// TwinCAT 3 PLC project PLC1
// ProgramVersion: 3.1.4024.0
// libraries:
//   Tc2_MC2, * (Beckhoff Automation GmbH)
//   Tc2_Standard, * (Beckhoff Automation GmbH)
//   Tc2_System, * (Beckhoff Automation GmbH)
//   Tc2_TcpIp, * (Beckhoff Automation GmbH)
//   Tc3_Module, * (Beckhoff Automation GmbH)
// project tree:
//   DUTs/ E_MelsecDevice.TcDUT, ST_MelsecSession.TcDUT, ST_QueuedCameraProduct.TcDUT, ST_Point2D.TcDUT, ST_QD75_Command.TcDUT, ST_QD75_Feedback.TcDUT
//   GVLs/ GVL_MD200_IO.TcGVL, GVL.TcGVL
//   / PlcTask.TcTTO
//   POUs/ FB_ConveyorEncoder.TcPOU, FB_ConveyorTracking4Pt.TcPOU, FB_InovanceMD200Conveyor.TcPOU, FB_EziServoControl.TcPOU, FB_MelsecEchoVerify.TcPOU, FB_MelsecDebugXY4Pt.TcPOU, FB_CameraProductQueue.TcPOU, FB_UpstreamCameraTracking4Pt.TcPOU, FB_XYTrackingManualAck.TcPOU, FB_MelsecRead.TcPOU, FB_MelsecTcpConfig.TcPOU, FB_MelsecWrite.TcPOU, FB_QD75CommandPublisher.TcPOU, MAIN.TcPOU
// real-time tasks:
//   TASK PlcTask: cycle T#10ms, priority 20, ADS port 350
// motion (NC):
//   TASK NC-Task 1 SAF: cycle T#2ms, priority 4, ADS port 501
//   TASK NC-Task 1 SVB: cycle T#10ms, priority 8, ADS port 511
//   AXIS Axis 1 (id 2)
//     General: UnitName=Degree
//     Velo: Maximum=50000
//     OtherSettings: AllowMotionCmdToSlave=true
//     encoder EncType=19
//       EncPara: ScaleFactorNumerator=360, ScaleFactorDenominator=10000, MaxCount=#xffffffff
//     drive DrvType=16
//       DrvPara: MaxCount=#xffffffff, DriveControlDWord=#x00020000
//         Analog: VeloReferenz=60000, TorqueSetpointScale=10, ScaleFactorActTorque=0.1
//         TimeComp: TaskDelayCycles=1
//     controller CtrType=1
//       CtrPara: PriorControlFactor=1
//         PosDiffControl: Range=60, Time=0.05
//         Observer: BandWidth=20
// I/O:
//   DEVICE Device 2 (EtherCAT), AmsNetId 10.81.27.140.3.1
//     Box 1 (NA-9286,Crevis) [NA-9286 EtherCAT Adapter, Crevis]
//       modules: Module 1 (ST-5101), Module 2 (ST-1228), Module 3 (ST-1228), Module 4 (ST-1228), Module 5 (ST-1228), Module 6 (ST-1228), Module 7 (ST-2318), Module 8 (ST-2318), Module 9 (ST-2318), Module 10 (ST-2318), Module 11 (ST-4424), Module 12 (ST-5114), Module 13 (ST-3214)
//     Drive 2 (Ezi-SERVO2 EtherCAT) [Ezi-SERVO2 EtherCAT]
// variable links:
//   NC-Task 1 SAF/Axes/Axis 1 <-> Device 2 (EtherCAT)/Drive 2 (Ezi-SERVO2 EtherCAT)
//     Drive/Inputs/In/nDcOutputTime <-> InfoData/DcOutputShift
//     Drive/Inputs/In/nState1 <-> CSP Inputs/Status Word
//     Drive/Inputs/In/nState2 <-> CSP Inputs/Status Word @bit 8
//     Drive/Inputs/In/nState4 @bit 1 <-> WcState/InputToggle
//     Drive/Inputs/In/nState4 <-> WcState/WcState
//     Drive/Outputs/Out/nCtrl1 <-> CSP Outputs/Control Word
//     Drive/Outputs/Out/nCtrl2 <-> CSP Outputs/Control Word @bit 8
//     Drive/Outputs/Out/nDataOut1 <-> CSP Outputs/Target Position
//     Enc/Inputs/In/nDataIn1 <-> CSP Inputs/Position Actual Value
//     Enc/Inputs/In/nDataIn3 <-> CSP Inputs/Touch probe 1 positive value
//     Enc/Inputs/In/nDataIn5 <-> CSP Inputs/Touch probe 2 positive value
//     Enc/Inputs/In/nDcInputTime <-> InfoData/DcInputShift
//     Enc/Inputs/In/nState4 @bit 1 <-> WcState/InputToggle
//     Enc/Inputs/In/nState4 <-> WcState/WcState
//     Enc/Inputs/In/nState5 <-> CSP Inputs/Touch probe status
//     Enc/Inputs/In/nState6 <-> CSP Inputs/Touch probe status @bit 8
//     Enc/Outputs/Out/nCtrl5 <-> CSP Outputs/Touch probe function
//     Enc/Outputs/Out/nCtrl6 <-> CSP Outputs/Touch probe function @bit 8
//   PLC1/PLC1 Instance <-> Device 2 (EtherCAT)/Box 1 (NA-9286,Crevis)
//     PlcTask Inputs/GVL.aIn[{0..15}] <-> Module 12 (ST-5114)/Input(s)/Byte {0..15}  (16 links)
//     PlcTask Inputs/GVL_MD200_IO.bEStopFeedback <-> Module 6 (ST-1228)/Input(s)/Byte 0
//     PlcTask Outputs/GVL.aOut[{0..3}] <-> Module 12 (ST-5114)/Output(s)/Byte {0..3}  (4 links)
//     PlcTask Outputs/GVL_MD200_IO.bRUN_DO <-> Module 10 (ST-2318)/Output(s)/Byte 0
//     PlcTask Outputs/GVL_MD200_IO.nAO1_Raw <-> Module 11 (ST-4424)/Output(s)/Analog Output Ch#1 Byte
//   PLC1/PLC1 Instance <-> NC-Task 1 SAF/Axes/Axis 1
//     PlcTask Inputs/MAIN.Axis1.NcToPlc <-> Outputs/ToPlc
//     PlcTask Outputs/MAIN.Axis1.PlcToNc <-> Inputs/FromPlc

CONFIGURATION PLC1
    RESOURCE PLC ON TwinCAT3
        TASK PlcTask(INTERVAL := T#10ms, PRIORITY := 20);
        PROGRAM MAIN WITH PlcTask : MAIN;
    END_RESOURCE
END_CONFIGURATION

// ---- DUTs/E_MelsecDevice.TcDUT
// Mã định danh vùng nhớ phần cứng Mitsubishi theo chuẩn MC Protocol Binary 3E Frame
TYPE E_MelsecDevice :
(
    DEV_D   := 16#A8, // Thanh ghi dữ liệu D (Data Register) - Word
    DEV_M   := 16#90, // Rơ-le nội bộ M (Internal Relay) - Bit / Word
    DEV_W   := 16#B4, // Thanh ghi liên kết W (Link Register) - Word
    DEV_R   := 16#AF, // Thanh ghi tệp R (File Register) - Word
    DEV_ZR  := 16#B0, // Thanh ghi tệp liên tục ZR (File Register Consecutive) - Word
    DEV_X   := 16#9C, // Ngõ vào vật lý X (Input) - Bit
    DEV_Y   := 16#9D, // Ngõ ra vật lý Y (Output) - Bit
    DEV_B   := 16#A0, // Rơ-le liên kết B (Link Relay) - Bit / Word
    DEV_L   := 16#92, // Rơ-le chốt L (Latch Relay) - Bit
    DEV_TN  := 16#C2, // Giá trị hiện tại Timer TN (Timer Current Value) - Word
    DEV_CN  := 16#C5  // Giá trị hiện tại Counter CN (Counter Current Value) - Word
);
END_TYPE

// ---- DUTs/ST_MelsecSession.TcDUT
TYPE ST_MelsecSession :
STRUCT
    hSocket     : T_HSOCKET; // Socket TCP dùng chung
    bConnected  : BOOL;      // TRUE khi đã kết nối PLC
    bBusy       : BOOL;      // TRUE khi Read hoặc Write đang giao dịch
    bError      : BOOL;      // Lỗi cuối cùng
    nErrorID    : UDINT;     // Mã lỗi cuối cùng
END_STRUCT
END_TYPE

// ---- DUTs/ST_QueuedCameraProduct.TcDUT
TYPE ST_QueuedCameraProduct :
STRUCT
    bValid                    : BOOL;
    nProductID                : UDINT;
    nState                    : INT; // 0 EMPTY, 1 WAIT_ROBOT, 2 GEOMETRIC_WINDOW
    bAllCornersInside         : BOOL;
    bForecastWindowOK         : BOOL;
    rEncoderAtExposure_mm     : LREAL;
    rCenterAtExposureX_mm     : LREAL;
    rCenterAtExposureY_mm     : LREAL;
    rThetaRobot_deg           : LREAL;
    rTravel_mm                : LREAL;
    rCenterNowX_mm            : LREAL;
    rCenterNowY_mm            : LREAL;
    aCornerBase               : ARRAY[1..4] OF ST_Point2D;
    aCornerNow                : ARRAY[1..4] OF ST_Point2D;
END_STRUCT
END_TYPE

// ---- DUTs/ST_Point2D.TcDUT
TYPE ST_Point2D :
STRUCT
    X : LREAL; // Tọa độ X (mm)
    Y : LREAL; // Tọa độ Y (mm)
END_STRUCT
END_TYPE

// ---- DUTs/ST_QD75_Command.TcDUT
TYPE ST_QD75_Command :
STRUCT
    Target_X       : DINT; // D100..D101: Tọa độ đón đầu trục X (0.1 um)
    Target_Y       : DINT; // D102..D103: Tọa độ trục Y đỉnh (0.1 um)
    Target_Z_Down  : DINT; // D104..D105: Độ cao hạ chấm keo (0.1 um, 4.0mm = 40000)
    Speed_Approach : DINT; // D106..D107: Vận tốc bay nội suy 3 trục (0.01 mm/min, 500mm/s = 3000000)
    Speed_Sync     : DINT; // D108..D109: Vận tốc đồng tốc trục X khi chấm keo (= V_conv * 6000)
    DeltaX_Sync    : DINT; // D110..D111: Quãng đường trượt đồng tốc 60ms (0.1 um)
    Target_Z_Safe  : DINT; // D112..D113: Độ cao an toàn khi rút kim (0.1 um, 0.0mm = 0)
    Vertex_Index   : INT;  // D114: Thứ tự đỉnh đang làm (1..4)
    Cmd_Start      : BOOL; // M1000: Kích chạy đỉnh đang nạp (TwinCAT -> PLC-Q)
END_STRUCT
END_TYPE

// ---- DUTs/ST_QD75_Feedback.TcDUT
TYPE ST_QD75_Feedback :
STRUCT
    Ack_Done    : BOOL; // M1001: PLC-Q báo Point 3 hoàn tất
    Robot_Busy  : BOOL; // M102: PLC-Q đang kiểm tra/nạp/chạy
    In_Position : BOOL; // M103: Đỉnh đã hoàn tất, chờ Master hạ M1000
    Robot_Alarm : BOOL; // M104: QD75 hoặc kiểm tra biên báo lỗi
END_STRUCT
END_TYPE

// ---- GVLs/GVL_MD200_IO.TcGVL
VAR_GLOBAL
    // E-stop circuit HEALTHY auxiliary contact feedback.
    // REVIEW BEFORE ACTIVATION: maps ST-1228 SLOT 6 / DI0 (physical terminal 0).
    // This is a PROPOSED wiring channel, not confirmed by cabinet visual inspection.
    // It must be wired to the healthy auxiliary feedback of an independent
    // hardwired emergency-stop safety circuit. TRUE = safety chain healthy.
    // This input alone is NOT an emergency-stop device.
    {attribute 'TcLinkToOSO' := '<0,1,0>TIID^Device 2 (EtherCAT)^Box 1 (NA-9286,Crevis)^Module 6 (ST-1228)^Input(s)^Byte 0'}
    bEStopFeedback AT %I* : BOOL := FALSE;

    // MD200 physical process-image channels, staged for deliberate link review.
    // ST-4424 Module 11 Channel AO1 (physical terminal 1, 0-10V).
    // UINT 16 bit with 12-bit useful range 0..4095.
    {attribute 'TcLinkTo' := 'TIID^Device 2 (EtherCAT)^Box 1 (NA-9286,Crevis)^Module 11 (ST-4424)^Output(s)^Analog Output Ch#1 Byte'}
    nAO1_Raw AT %Q* : UINT := 0;

    // Staged logical RUN: ST-2318 Module 10 immediately before AO module.
    // DO0 is bit 0 of Output(s)^Byte 0; map ONLY one bit (not entire BYTE).
    // WARNING: physical DO0/pin 0 must be confirmed unused and NPN wiring
    // checked by the on-site technician BEFORE activating this configuration.
    // All runtime software permits remain FALSE by default.
    {attribute 'TcLinkToOSO' := '<0,1,0>TIID^Device 2 (EtherCAT)^Box 1 (NA-9286,Crevis)^Module 10 (ST-2318)^Output(s)^Byte 0'}
    bRUN_DO AT %Q* : BOOL := FALSE;
END_VAR

// ---- GVLs/GVL.TcGVL
VAR_GLOBAL
    aIn  AT %I* : ARRAY[0..15] OF BYTE;  // TxPDO 16 byte
    aOut AT %Q* : ARRAY[0..3]  OF BYTE;  // RxPDO 4 byte
END_VAR

// ---- POUs/MAIN.TcPOU
PROGRAM MAIN
VAR
    // ================================================================
    // 1. KẾT NỐI TCP VỚI CPU MITSUBISHI Q06UDEH (CỔNG 5010)
    // ================================================================
    stMelsec            : ST_MelsecSession; // Session TCP dùng chung
    fbMelsecConfig      : FB_MelsecTcpConfig;

    bTcpEnable          : BOOL := TRUE;     // Tự động kết nối và duy trì kết nối mạng
    sPlcQ_IP            : STRING(15) := '192.168.3.39'; // IP của PLC-Q
    nPlcQ_Port          : UDINT := 5010;   // Cổng Port MC Protocol 5010

    bPlcQConnected      : BOOL;             // ĐÈN BÁO: TRUE = Đã thông mạng với PLC-Q
    bPlcQError          : BOOL;
    nPlcQErrorID        : UDINT;

    // ================================================================
    // 2. TEST TRUYỀN THÔNG THỦ CÔNG SANG PLC-Q (KHI bStartGlueCycle = FALSE)
    // ================================================================
    bTest_WriteD100     : BOOL := FALSE;    // Click đúp TRUE -> Ghi nTest_D100_Val vào D100-D101
    nTest_D100_Val      : DINT := 100;      // Số 32-bit gửi thử sang D100
    bTest_WriteM1000    : BOOL := FALSE;    // Click đúp TRUE -> Ghi bit M1000
    bTest_M1000_Val     : BOOL := TRUE;     // Giá trị bit M1000 muốn ghi (TRUE=ON, FALSE=OFF)
    bTest_ReadM1001     : BOOL := FALSE;    // Click đúp TRUE -> Đọc bit M1001 từ PLC-Q
    bTest_M1001_Result  : BOOL;             // Giá trị M1001 đọc được từ PLC-Q

    // ================================================================
    // 3. ENCODER BĂNG TẢI: ST-5114 MODULE 12
    // ================================================================
    fbConveyor          : FB_ConveyorEncoder;

    nEncoderPulse       : UINT;            // HARDWARE RAW counter, NOT zeroed on TwinCAT boot
    nEncoderPulseSinceStart : DINT := 0; // VIRTUAL count starting from 0 on PLC boot
    nEncoderDelta       : INT;             // Xung thay đổi trong 10 ms
    rConveyorSpeed      : LREAL;           // Vận tốc băng tải lọc mượt, mm/s
    rConveyorSpeedMPM   : LREAL;           // Vận tốc băng tải, m/phút
    rConveyorDist       : LREAL;           // Tổng quãng đường băng tải, mm

    // ================================================================
    // ================================================================
    // MD200 VFD PREPARATION / VIRTUAL ONLY (NO PHYSICAL I/O MAPPING).
    // Outputs remain disconnected from Crevis ST-2318 and ST-4424.
    // ================================================================
    fbMD200_VFD               : FB_InovanceMD200Conveyor;
    // Global normal-PLC motion inhibit, NOT an emergency stop safety function.
    // TRUE only when the auxiliary feedback from hardwired EStop is healthy.
    bSystemEStopOK             : BOOL := FALSE;
    bSystemStopRequested       : BOOL := TRUE;
    // Only 3 operator-visible MD200 signals: EStopOK monitor, START and Hz.
    // EStopOK is derived from the wired digital feedback, NOT an HMI override.
    bMD200_EStopOK           : BOOL := FALSE;
    bMD200_Start             : BOOL := FALSE;
    rMD200_SetFrequency_Hz    : LREAL := 0.0;
    // Diagnostics (read-only outputs from the FB)
    bMD200_DO_RunVirtual      : BOOL;
    nMD200_AO_RawVirtual      : INT;
    rMD200_AO_VoltsVirtual    : LREAL;
    rMD200_Target_Hz          : LREAL;
    rMD200_Ramped_Hz          : LREAL;
    bMD200_AtTarget           : BOOL;
    bMD200_Limited            : BOOL;
    nMD200_Status             : UINT;

    // ================================================================
    // 4. EZI-SERVO: TRỤC QUAY ĐƠN VỊ DEGREE
    // ================================================================
    Axis1               : AXIS_REF;

    fbServo             : FB_EziServoControl;

    bServo_Enable       : BOOL := FALSE;     // TRUE = Servo ON / giữ cốt
    bServo_Reset        : BOOL := FALSE;    // TRUE một chu kỳ = Reset Alarm
    bServo_JogFwd       : BOOL := FALSE;    // TRUE = chạy thuận
    bServo_JogBwd       : BOOL := FALSE;    // TRUE = chạy nghịch

    rServo_Speed        : LREAL := 100.0;   // Degree/s
    rServo_Acc          : LREAL := 400.0;   // Degree/s2
    rServo_Dec          : LREAL := 400.0;   // Degree/s2

    bServo_Ready        : BOOL;             // TRUE = Servo ON
    rServo_ActPos_Deg   : LREAL;            // Góc thực tế, Degree
    rServo_ActVel_Deg_s : LREAL;            // Vận tốc thực tế, Degree/s

    // ================================================================
    // 5. TRACKING 4 ĐIỂM: CAMERA + ENCODER
    // ================================================================
    fbTracking4Pt       : FB_ConveyorTracking4Pt;

    bSystemReset        : BOOL := FALSE;    // TRUE một chu kỳ: reset mốc phần mềm về 0
    // Camera giả lập test
    bCameraTrigger      : BOOL := FALSE;    // FALSE -> TRUE: chốt sản phẩm mới
    rCameraCenterX      : LREAL := 0.0;     // Camera input, starts 0 until REAL result
    rCameraCenterY      : LREAL := 0.0;     // Camera input, starts 0 until REAL result
    rCameraAngleDeg     : LREAL := 0.0;     // Góc phôi, Degree
    rProductLength      : LREAL := 40.0;    // mm
    rProductWidth       : LREAL := 40.0;    // mm

    // Kết quả debug Tracking
    bProductValid       : BOOL;
    nPulseAtCamera      : UINT;
    nPulseTravel        : INT;
    rPartTravel_mm      : LREAL;

    aCornerBase         : ARRAY[1..4] OF ST_Point2D;
    aCornerNow          : ARRAY[1..4] OF ST_Point2D;

    // ================================================================
    // 6. QD75 COMMAND PUBLISHER: ĐIỀU PHỐI 4 ĐỈNH SANG PLC-Q
    // ================================================================
    fbPublisher         : FB_QD75CommandPublisher;

    // ================================================================
    // AUTO DISPATCH: opt-in only, requires an actual camera event.
    // No motor/robot command can be emitted by this feature by default.
    // ================================================================
    bAutoDispatchEnable : BOOL := FALSE;   // Operator enables auto sequence only after commissioning
    bAutoDispatchArm    : BOOL := FALSE;   // Independent arm interlock
    fbAutoCameraEdge    : R_TRIG;
    tonAutoProductTTL   : TON;
    bAutoPendingProduct : BOOL := FALSE;
    bAutoStartPulse     : BOOL := FALSE;
    nAutoDispatchState  : INT := 0;       // 0 idle, 1 queued, 2 speed invalid, 3 TCP busy/offline, 4 motion busy, 5 expired, 6 invalid product, 10 request issued
    nAutoStartRequests  : UDINT := 0;

    // ================================================================
    // 6A. ISOLATED DATA-ONLY XY DEBUG (D100-D103 + D114, NO Z/M1000)
    // Requires physically stopped conveyor and robot; service opt-in.
    // ================================================================
    fbDebugXY           : FB_MelsecDebugXY4Pt;
    bDebugXYPermit      : BOOL := FALSE; // Set TRUE only during maintenance
    bDebugXYExecute     : BOOL := FALSE; // Pulse FALSE -> TRUE once
    bDebugXYAbort       : BOOL := FALSE;
    rDebugCenterX       : LREAL := 50.0;
    rDebugCenterY       : LREAL := 85.0;
    rDebugAngleDeg      : LREAL := 0.0;
    rDebugLength        : LREAL := 40.0;
    rDebugWidth         : LREAL := 40.0;
    bDebugXYMachineStopped : BOOL;
    bDebugXYBusy        : BOOL;
    bDebugXYDone        : BOOL; // Data ACK only, not robot done
    bDebugXYError       : BOOL;
    nDebugXYErrorCode   : INT;
    nDebugXYCommError   : UDINT;
    nDebugXYState       : INT;
    nDebugXYVertex      : INT;
    nDebugXYPassed      : INT;
    nDebugXYWriteX      : DINT;
    nDebugXYWriteY      : DINT;
    nDebugXYReadX       : DINT;
    nDebugXYReadY       : DINT;
    nDebugXYReadVertex  : UINT;
    bDebugXYReadbackOK  : BOOL;
    bDebugXYAllBitsLow  : BOOL;
    bDebugXYRestored    : BOOL;

    // ================================================================
    // UPSTREAM CAMERA -> ENCODER -> ROBOT XY
    // Camera provides CENTER X/Y (physical mm) and ANGLE, not corners.
    // Calibration and real camera transport MUST be proven before enabling.
    // ================================================================
    fbUpstreamTrack      : FB_UpstreamCameraTracking4Pt;
    bUpstreamReset       : BOOL := FALSE;
    bCameraExposeTrigger : BOOL := FALSE; // Pulse from strobe/trigger at IMAGE exposure
    fbCameraExposeEdge   : R_TRIG;
    fbVisionResultEdge   : R_TRIG;
    tonExposureTTL       : TON;
    bExposureEncoderLatched : BOOL := FALSE;
    rEncoderAtExposure_mm   : LREAL := 0.0;
    bVisionFeedVerified  : BOOL := FALSE; // FALSE until actual camera bridge is installed
    bVisionCalibrationOK : BOOL := FALSE; // TRUE only after physical frame calibration
    rCameraToWorkStart_mm : LREAL := 0.0; // USER-EDITABLE POSITIVE DISTANCE (mm); 0 blocks tracking
    rCamToRobotX_mm      : LREAL := 0.0;  // Fine X offset after measuring camera-to-work distance
    rCamToRobotY_mm      : LREAL := 0.0;
    rCamToRobotYaw_deg   : LREAL := 0.0;
    bUpstreamCaptured    : BOOL;
    bUpstreamInWorkspace : BOOL;
    bUpstreamPastRobot   : BOOL;
    nUpstreamError       : INT;
    rUpstreamDrift_mm    : LREAL;
    rUpstreamCenterX     : LREAL;
    rUpstreamCenterY     : LREAL;
    rUpstreamNowX        : LREAL;
    rUpstreamNowY        : LREAL;
    rToRobotWorkStart_mm : LREAL; // Countdown to X=0, 0 after entering
    aUpstreamCornerNow   : ARRAY[1..4] OF ST_Point2D;

    // ================================================================
    // CAMERA FIFO MONITOR (DATA ONLY): independent 8-product queue.
    // Camera returns CENTER X/Y in mm and ANGLE in degrees, NOT corners.
    // No robot Publisher connection or M1000 writes in this stage.
    // ================================================================
    fbCameraQueue        : FB_CameraProductQueue;
    bLegacyMotionPublisherAllow : BOOL := FALSE; // explicit safety gate: NO robot in FIFO stage
    bQueueReset          : BOOL := FALSE;
    bQueueSimMode        : BOOL := FALSE; // explicit dry-run mode only
    bQueueSimExposure    : BOOL := FALSE;
    bQueueSimResult      : BOOL := FALSE;
    bQueueSimCompleteHead : BOOL := FALSE; // virtual DONE, NOT Mitsubishi ACK
    nQueueCount          : INT;
    nQueueHeadProductID  : UDINT;
    nQueueHeadState      : INT;
    bQueueHeadValid      : BOOL;
    bQueueHeadAllInside  : BOOL; // geometric observation only
    bQueueHeadForecastOK : BOOL; // theoretical estimate, NOT permission to move
    rQueueHeadTravel_mm  : LREAL;
    rQueueToWorkStart_mm : LREAL;
    rQueueHeadX_mm       : LREAL;
    rQueueHeadY_mm       : LREAL;
    aQueueHeadCornerNow  : ARRAY[1..4] OF ST_Point2D;
    nQueueAccepted       : UDINT;
    nQueueRejected       : UDINT;
    nQueueMissed         : UDINT;
    nQueueSimCompleted   : UDINT;
    bQueueInputFault     : BOOL;
    nQueueErrorCode      : INT;

    // ================================================================
    // MANUAL ACK BENCH MODE ONLY: no M1000, Z, QD75 or valve writes.
    // User reserves/audits a spare PLC bit (proposed M2100), NOT M1001.
    // ================================================================
    fbXYManualAck        : FB_XYTrackingManualAck;
    bXYManualPermit      : BOOL := FALSE;
    bXYManualExecute     : BOOL := FALSE;
    bXYManualAbort       : BOOL := FALSE;
    bXYManualAckBitAudited : BOOL := FALSE;
    nXYManualAckMAddress : UDINT := 2100;
    bXYManualSafe        : BOOL;
    bXYManualBusy        : BOOL;
    bXYManualDone        : BOOL;
    bXYManualError       : BOOL;
    bXYManualRestored    : BOOL;
    nXYManualErrorCode   : INT;
    nXYManualCommError   : UDINT;
    nXYManualState       : INT;
    nXYManualVertex      : INT;
    nXYManualAcked       : INT;
    nXYManualSentX       : DINT;
    nXYManualSentY       : DINT;
    nXYManualReadX       : DINT;
    nXYManualReadY       : DINT;
    nXYManualReadVertex  : UINT;
    bXYManualReadbackOK  : BOOL;

    // Lệnh chu trình chấm keo
    bStartGlueCycle     : BOOL := FALSE;   // FALSE -> TRUE: kích chạy chu trình 4 đỉnh
    bGlueResetFault     : BOOL := FALSE;    // Operator acknowledges latched fault
    bEnableManualWrite  : BOOL := FALSE;    // OFF unless supervised maintenance
    bAbortGlueCycle     : BOOL := FALSE;   // TRUE: dừng khẩn cấp (ghi M105)

    // Trạng thái giám sát chu trình
    bGlueCycleBusy      : BOOL;            // Đang chạy 4 đỉnh
    bGlueCycleDone      : BOOL;            // Hoàn tất cả 4 đỉnh
    bGlueCycleError     : BOOL;            // Báo lỗi
    bStopCommandConfirmed : BOOL;          // PLC đã xác nhận 2 lệnh dừng qua TCP
    nGlueCurVertex      : INT;             // Đỉnh đang thực hiện (1..4)
    nGlueCommErrorID    : UDINT;           // raw error from MC socket or Mitsubishi
    nGlueErrorCode      : INT;             // Mã lỗi (501..503, 900..921)

    // ================================================================
    // 7. MC 3E TCP WORD/BIT ECHO VERIFY (OFF by default)
    //    Explicit permission required. Never use motion/handshake addresses.
    // ================================================================
    fbEchoWord          : FB_MelsecEchoVerify;
    fbEchoBit           : FB_MelsecEchoVerify;
    bEchoPermit         : BOOL := FALSE;    // Maintenance only
    bEchoMachineSafe    : BOOL := FALSE;    // Operator confirmed gantry safe
    bEchoAddressChecked : BOOL := FALSE;    // Both addresses audited in PLC/HMI
    bEchoRequestWord    : BOOL := FALSE;    // One-shot rising edge
    bEchoRequestBit     : BOOL := FALSE;    // One-shot rising edge
    nEchoDAddress       : UDINT := 0;       // Must be an approved unused D>=3000
    nEchoMAddress       : UDINT := 0;       // Must be an approved unused M>=2000
    wEchoTestValue      : WORD := 16#A55A;
    bEchoTestValue      : BOOL := TRUE;
    bEchoWordDone       : BOOL;
    bEchoWordBusy       : BOOL;
    bEchoWordError      : BOOL;
    bEchoWordMatch      : BOOL;
    bEchoWordRestored   : BOOL;
    bEchoWordRestoreUncertain : BOOL;
    nEchoWordErrorID    : UDINT;
    wEchoWordBefore     : WORD;
    wEchoWordAfter      : WORD;
    bEchoBitDone        : BOOL;
    bEchoBitBusy        : BOOL;
    bEchoBitError       : BOOL;
    bEchoBitMatch       : BOOL;
    bEchoBitRestored    : BOOL;
    bEchoBitRestoreUncertain : BOOL;
    nEchoBitErrorID     : UDINT;
    bEchoBitBefore      : BOOL;
    bEchoBitAfter       : BOOL;
END_VAR

// ================================================================
// 1. TCP CONFIG: Kết nối / tự reconnect đến PLC-Q
// ================================================================
fbMelsecConfig(
    bEnable     := bTcpEnable,
    sRemoteHost := sPlcQ_IP,
    nRemotePort := nPlcQ_Port,
    stSession   := stMelsec
);

// Biến trạng thái đưa ra ngoài để Online debug dễ
bPlcQConnected := stMelsec.bConnected;
bPlcQError     := stMelsec.bError;
nPlcQErrorID   := stMelsec.nErrorID;

// ================================================================
// SYSTEM-WIDE NORMAL PLC INTERLOCK FROM ONE PHYSICAL E-STOP FEEDBACK.
// NOT SAFETY RATED. Hardware chain must remove hazardous motion in both
// MD200 and Mitsubishi QD75 independently of TwinCAT and Ethernet.
// HMI/ADS must NOT force this input. Keep network alive for best-effort
// Q-PLC cancel. Clear old command bits to prevent unintended restart.
// ================================================================
bSystemEStopOK := GVL_MD200_IO.bEStopFeedback;
bSystemStopRequested := NOT bSystemEStopOK;
IF bSystemStopRequested THEN
    bMD200_Start := FALSE;
    bServo_Enable := FALSE;
    bServo_JogFwd := FALSE;
    bServo_JogBwd := FALSE;
    bServo_Reset := FALSE;
    bStartGlueCycle := FALSE;
    bAutoDispatchEnable := FALSE;
    bAutoDispatchArm := FALSE;
    bAutoPendingProduct := FALSE;
    bAutoStartPulse := FALSE;
    bLegacyMotionPublisherAllow := FALSE;
    bEnableManualWrite := FALSE;
    bTest_WriteM1000 := FALSE;
    bTest_WriteD100 := FALSE;
    bDebugXYPermit := FALSE;
    bDebugXYExecute := FALSE;
    bXYManualPermit := FALSE;
    bXYManualExecute := FALSE;
    bEchoPermit := FALSE;
    bEchoRequestWord := FALSE;
    bEchoRequestBit := FALSE;
    bQueueSimMode := FALSE;
END_IF;


// ================================================================
// 2. ENCODER BĂNG TẢI: ST-5114 INPUT BYTE 0 + BYTE 1
// ================================================================
fbConveyor(
    bByte0          := GVL.aIn[0],
    bByte1          := GVL.aIn[1],
    rK_mm           := 0.476475,
    rCycleTime      := 0.01,

    nRawPulse       => nEncoderPulse,
    nDeltaPulse     => nEncoderDelta,
    rSpeed_mm_s     => rConveyorSpeed,
    rSpeed_m_min    => rConveyorSpeedMPM,
    rTotalDist_mm   => rConveyorDist
);

// The display count starts at 0 on PLC boot, unlike nEncoderPulse,
// which is the actual hardware ST-5114 counter and may be non-zero.
// DINT is used to avoid modulo-65536 wrap in this visual counter.
nEncoderPulseSinceStart := nEncoderPulseSinceStart + INT_TO_DINT(nEncoderDelta);

// ================================================================
// ================================================================
// MD200 SIMPLE: EStop feedback, START request, 0..25Hz only.
// Actual emergency stop MUST act independently through the hardwired
// safety circuit. Software feedback is a monitor, not a safety device.
// ================================================================
bMD200_EStopOK := bSystemEStopOK;
fbMD200_VFD(
    bEStopOK            := bMD200_EStopOK,
    bStart              := bMD200_Start,
    rFrequencySet_Hz    := rMD200_SetFrequency_Hz,
    bDO_RunForward      => bMD200_DO_RunVirtual,
    nAO_12bitRaw        => nMD200_AO_RawVirtual,
    rAO_Volts           => rMD200_AO_VoltsVirtual,
    rTarget_Hz          => rMD200_Target_Hz,
    rRamped_Hz          => rMD200_Ramped_Hz,
    bAtTarget           => bMD200_AtTarget,
    bLimited25Hz        => bMD200_Limited,
    nStatus             => nMD200_Status
);

// Only ONE producer writes process-image outputs; no direct ADS test signal.
// FB implements 25Hz clamp and all software/verified interlock checks.
// In this isolated stage the outputs are AT %Q* process tags, still
// NOT linked to physical Crevis channels until I/O link verification.
IF (nMD200_AO_RawVirtual >= 0) AND (nMD200_AO_RawVirtual <= 4095) THEN
    GVL_MD200_IO.nAO1_Raw := INT_TO_UINT(nMD200_AO_RawVirtual);
ELSE
    GVL_MD200_IO.nAO1_Raw := 0;
END_IF;
GVL_MD200_IO.bRUN_DO := bMD200_DO_RunVirtual;

// ================================================================
// 3. EZI-SERVO: ENABLE, RESET, JOG VÀ GIÁM SÁT
// ================================================================
fbServo(
    Axis            := Axis1,
    bEnable         := bServo_Enable AND bSystemEStopOK,
    bResetFault     := bServo_Reset AND bSystemEStopOK,
    bJogFwd         := bServo_JogFwd AND bSystemEStopOK,
    bJogBwd         := bServo_JogBwd AND bSystemEStopOK,
    rTargetVelocity := rServo_Speed,
    rAcc            := rServo_Acc,
    rDec            := rServo_Dec,

    bReady          => bServo_Ready,
    rActPos_Deg     => rServo_ActPos_Deg,
    rActVel_Deg     => rServo_ActVel_Deg_s
);

IF bServo_Reset THEN
    bServo_Reset := FALSE;
END_IF;


// ================================================================
// 4. TRACKING 4 ĐIỂM: CAMERA + ENCODER
// ================================================================
fbTracking4Pt(
    bResetSystem   := bSystemReset OR bSystemStopRequested,
    bCameraResult  := FALSE, // legacy tracker intentionally disconnected from Camera
    bAcceptCamera  := FALSE, // all live products must use FIFO, not legacy single item
    rCenterX_mm    := rCameraCenterX,
    rCenterY_mm    := rCameraCenterY,
    rAngleDeg      := rCameraAngleDeg,
    rLength_mm     := rProductLength,
    rWidth_mm      := rProductWidth,

    nEncoderNow    := nEncoderPulse,
    rMmPerPulse    := 0.476475,
    rXMaxLimit_mm  := 180.0,

    bProductValid  => bProductValid,
    nPulseAtCamera => nPulseAtCamera,
    nPulseTravel   => nPulseTravel,
    rTravel_mm     => rPartTravel_mm,
    aCornerBase    => aCornerBase,
    aCornerNow     => aCornerNow
);

IF bSystemReset THEN
    bSystemReset := FALSE;
END_IF;

// ================================================================
// 4A. CAMERA -> AUTO DISPATCH (explicitly DISABLED until commissioned)
// The camera event queues one product. No command is sent merely
// because bProductValid remains TRUE from a previous snapshot.
// ================================================================
fbAutoCameraEdge(CLK := bCameraTrigger);
bAutoStartPulse := FALSE;

// A pending camera event has a bounded lifetime (no stale product commands).
tonAutoProductTTL(IN := bAutoPendingProduct, PT := T#750MS);

IF bSystemStopRequested OR NOT bAutoDispatchEnable OR NOT bAutoDispatchArm OR bAbortGlueCycle
   OR bGlueResetFault OR bGlueCycleError OR bEchoPermit OR bDebugXYPermit OR bXYManualPermit THEN
    bAutoPendingProduct := FALSE;
    nAutoDispatchState := 0;
ELSIF fbAutoCameraEdge.Q AND bProductValid AND NOT bGlueCycleBusy THEN
    bAutoPendingProduct := TRUE;
    nAutoDispatchState := 1;
END_IF;

IF bAutoPendingProduct THEN
    IF tonAutoProductTTL.Q THEN
        bAutoPendingProduct := FALSE;
        nAutoDispatchState := 5; // Stale camera event discarded
    ELSIF NOT bProductValid THEN
        bAutoPendingProduct := FALSE;
        nAutoDispatchState := 6;
    ELSIF (rConveyorSpeed <= 0.0) OR (rConveyorSpeed > 1000.0) THEN
        nAutoDispatchState := 2; // Invalid conveyor speed; do not write 0 speed to QD75
    ELSIF NOT bPlcQConnected OR stMelsec.bBusy THEN
        nAutoDispatchState := 3;
    ELSIF bGlueCycleBusy OR bStartGlueCycle OR bEnableManualWrite
        OR bEchoWordBusy OR bEchoBitBusy THEN
        nAutoDispatchState := 4;
    ELSE
        bAutoStartPulse := TRUE; // Exactly one scan; Publisher performs PLC preflight
        bAutoPendingProduct := FALSE;
        nAutoStartRequests := nAutoStartRequests + 1;
        nAutoDispatchState := 10;
    END_IF;
END_IF;


// ================================================================
// 5. QD75 COMMAND PUBLISHER: ĐIỀU PHỐI 4 ĐỈNH & TEST THỦ CÔNG
// ================================================================
fbPublisher(
    stSession           := stMelsec,
    bStartCycle         := (bStartGlueCycle OR bAutoStartPulse) AND bSystemEStopOK AND bLegacyMotionPublisherAllow AND NOT bQueueSimMode AND NOT bEchoPermit AND NOT bEchoWordBusy AND NOT bEchoBitBusy AND NOT bDebugXYPermit AND NOT bDebugXYBusy AND NOT bXYManualPermit AND NOT bXYManualBusy,
    // Best-effort TCP cancellation only; cannot replace independent QD75
    // hardwired EStop. Avoid sending M105 when publisher is idle.
    bAbortCycle         := bAbortGlueCycle OR
                           (bSystemStopRequested AND
                             (bGlueCycleBusy OR (fbPublisher.nState = 70)
                              OR (fbPublisher.nState = 95))),
    bProductValid       := bProductValid,
    rEncoderDist_mm     := rConveyorDist,
    bResetFault         := bGlueResetFault AND bSystemEStopOK,
    bEnableManualWrite  := bEnableManualWrite AND bSystemEStopOK AND NOT bDebugXYPermit AND NOT bXYManualPermit,

    // Tọa độ 4 góc thời gian thực từ khối Tracking
    aCornerNow          := aCornerNow,
    rConveyorSpeed_mm_s := rConveyorSpeed,

    // Động học
    rFlyTime_s          := 0.120,
    rApproachSpeed_mm_s := 500.0,
    rSyncTime_s         := 0.060,
    rZDown_mm           := 4.0,
    rZSafe_mm           := 0.0,

    // Chế độ test thủ công (chỉ có tác dụng khi bStartGlueCycle = FALSE)
    bManualWriteD100    := bTest_WriteD100 AND bSystemEStopOK AND bLegacyMotionPublisherAllow AND NOT bQueueSimMode AND NOT bDebugXYPermit AND NOT bXYManualPermit,
    nD100_ManualVal     := nTest_D100_Val,
    bManualWriteM1000   := bTest_WriteM1000 AND bSystemEStopOK AND bLegacyMotionPublisherAllow AND NOT bQueueSimMode AND NOT bDebugXYPermit AND NOT bXYManualPermit,
    bM1000_ManualVal    := bTest_M1000_Val,
    bManualReadM1001    := bTest_ReadM1001 AND bSystemEStopOK AND NOT bDebugXYPermit AND NOT bXYManualPermit,

    // Giám sát
    bBusy               => bGlueCycleBusy,
    bDone               => bGlueCycleDone,
    bError              => bGlueCycleError,
    nErrorCode          => nGlueErrorCode,
    nLastCommError      => nGlueCommErrorID,
    nCurrentVertex      => nGlueCurVertex,
    bM1001_ReadBack     => bTest_M1001_Result,
    bStopCommandConfirmed => bStopCommandConfirmed
);

// Tự động nhả cờ kích test sau khi lệnh được nhận
IF bTest_WriteD100 AND NOT fbPublisher.bManualWriteD100 THEN
    bTest_WriteD100 := FALSE;
END_IF;

IF bTest_WriteM1000 AND NOT fbPublisher.bManualWriteM1000 THEN
    bTest_WriteM1000 := FALSE;
END_IF;

IF bTest_ReadM1001 AND NOT fbPublisher.bManualReadM1001 THEN
    bTest_ReadM1001 := FALSE;
END_IF;

// ================================================================
// 6. OPTIONAL WRITE -> READ SAME ADDRESS -> RESTORE -> VERIFY.
//    Never activated automatically. Does not touch motion D100/M1000.
//    Only one echo request at a time; uses shared stSession mutex.
// ================================================================
fbEchoWord(
    stSession := stMelsec,
    bExecute := bEchoRequestWord AND bSystemEStopOK AND NOT bEchoRequestBit,
    bEnable := bEchoPermit AND bSystemEStopOK AND NOT bGlueCycleBusy AND NOT bStartGlueCycle
               AND NOT bEnableManualWrite AND NOT bEchoBitBusy AND NOT bDebugXYPermit AND NOT bXYManualPermit,
    bAddressVerifiedUnused := bEchoAddressChecked,
    bMachineSafe := bEchoMachineSafe,
    bBitDevice := FALSE,
    nAddress := nEchoDAddress,
    wTestValue := wEchoTestValue,
    bBusy => bEchoWordBusy,
    bDone => bEchoWordDone,
    bError => bEchoWordError,
    bMatch => bEchoWordMatch,
    bRestored => bEchoWordRestored,
    bRestoreUncertain => bEchoWordRestoreUncertain,
    nErrorID => nEchoWordErrorID,
    wOriginal => wEchoWordBefore,
    wReadBack => wEchoWordAfter
);

fbEchoBit(
    stSession := stMelsec,
    bExecute := bEchoRequestBit AND bSystemEStopOK AND NOT bEchoRequestWord,
    bEnable := bEchoPermit AND bSystemEStopOK AND NOT bGlueCycleBusy AND NOT bStartGlueCycle
               AND NOT bEnableManualWrite AND NOT bEchoWordBusy AND NOT bDebugXYPermit AND NOT bXYManualPermit,
    bAddressVerifiedUnused := bEchoAddressChecked,
    bMachineSafe := bEchoMachineSafe,
    bBitDevice := TRUE,
    nAddress := nEchoMAddress,
    bTestValue := bEchoTestValue,
    bBusy => bEchoBitBusy,
    bDone => bEchoBitDone,
    bError => bEchoBitError,
    bMatch => bEchoBitMatch,
    bRestored => bEchoBitRestored,
    bRestoreUncertain => bEchoBitRestoreUncertain,
    nErrorID => nEchoBitErrorID,
    bOriginal => bEchoBitBefore,
    bReadBack => bEchoBitAfter
);

// ================================================================
// 7. DATA-ONLY DIAGNOSTIC: REAL TwinCAT -> MC TCP -> Mitsubishi.
// Operator must stop servo/conveyor, and provide two rising-edge
// flags (Permit=TRUE, Execute pulse). No Z, speed, M1000 or Y writes.
// ================================================================
bDebugXYMachineStopped :=
    NOT bServo_JogFwd AND NOT bServo_JogBwd
    AND (ABS(rServo_ActVel_Deg_s) < 0.2)
    AND (ABS(rConveyorSpeed) < 0.5)
    AND NOT bGlueCycleBusy AND NOT bStartGlueCycle
    AND NOT bAbortGlueCycle AND NOT bGlueCycleError;

fbDebugXY(
    stSession := stMelsec,
    bExecute := bDebugXYExecute AND bSystemEStopOK,
    bPermit := bDebugXYPermit AND bSystemEStopOK AND NOT bXYManualPermit AND NOT bEchoPermit
               AND NOT bEnableManualWrite AND NOT bAutoDispatchEnable
               AND NOT bAutoDispatchArm,
    bMachineStopped := bDebugXYMachineStopped,
    bPublisherIdle := (fbPublisher.nState = 0)
                      AND NOT bEchoWordBusy AND NOT bEchoBitBusy
                      AND NOT bTest_WriteM1000 AND NOT bTest_WriteD100,
    bAbort := bDebugXYAbort OR bSystemStopRequested,
    rCenterX_mm := rDebugCenterX,
    rCenterY_mm := rDebugCenterY,
    rAngleDeg := rDebugAngleDeg,
    rLength_mm := rDebugLength,
    rWidth_mm := rDebugWidth,
    tHold := T#10S,
    bBusy => bDebugXYBusy,
    bDone => bDebugXYDone,
    bError => bDebugXYError,
    nErrorCode => nDebugXYErrorCode,
    nCommErrorID => nDebugXYCommError,
    nState => nDebugXYState,
    nCurrentVertex => nDebugXYVertex,
    nPassedVertices => nDebugXYPassed,
    nWriteX => nDebugXYWriteX,
    nWriteY => nDebugXYWriteY,
    nReadX => nDebugXYReadX,
    nReadY => nDebugXYReadY,
    nReadVertex => nDebugXYReadVertex,
    bLastReadbackOK => bDebugXYReadbackOK,
    bAllMotionBitsLow => bDebugXYAllBitsLow,
    bOriginalRestored => bDebugXYRestored
);

// ================================================================
// 8. TRACK CAMERA CENTER+ANGLE (mm) FROM UPSTREAM STATION.
// Image exposure precedes Camera processing result. Encoder must be
// latched at exposure event, not at the delayed result arrival.
// ================================================================
fbCameraExposeEdge(CLK := bCameraExposeTrigger);
IF fbCameraExposeEdge.Q AND bVisionFeedVerified THEN
    rEncoderAtExposure_mm := rConveyorDist;
    bExposureEncoderLatched := TRUE;
END_IF;
tonExposureTTL(IN := bExposureEncoderLatched, PT := T#5S);
IF tonExposureTTL.Q THEN
    bExposureEncoderLatched := FALSE; // Reject stale camera processing events
END_IF;
fbVisionResultEdge(CLK := bCameraTrigger AND bVisionFeedVerified);

fbUpstreamTrack(
    bReset := bUpstreamReset OR bSystemStopRequested,
    bCameraResult := bCameraTrigger AND bVisionFeedVerified AND bSystemEStopOK,
    bAcceptCamera := bSystemEStopOK AND NOT bXYManualBusy AND NOT bGlueCycleBusy AND NOT bDebugXYBusy,
    bCalibrationConfirmed := bVisionCalibrationOK AND bVisionFeedVerified,
    bExposureEncoderValid := bExposureEncoderLatched,
    rEncoderAtExposure_mm := rEncoderAtExposure_mm,
    rCameraCenterX_mm := rCameraCenterX,
    rCameraCenterY_mm := rCameraCenterY,
    rCameraAngleDeg := rCameraAngleDeg,
    rCameraToWorkStart_mm := rCameraToWorkStart_mm,
    rCameraToRobotX_mm := rCamToRobotX_mm,
    rCameraToRobotY_mm := rCamToRobotY_mm,
    rCameraToRobotYawDeg := rCamToRobotYaw_deg,
    rEncoderTotalDist_mm := rConveyorDist,
    rLength_mm := rProductLength,
    rWidth_mm := rProductWidth,
    rRobotXMin_mm := 0.0,
    rRobotXMax_mm := 180.0,
    rRobotYMin_mm := 0.0,
    rRobotYMax_mm := 170.0,
    bCaptured => bUpstreamCaptured,
    bInRobotWorkspace => bUpstreamInWorkspace,
    bAllCornersPastRobot => bUpstreamPastRobot,
    nErrorCode => nUpstreamError,
    rEncoderTravel_mm => rUpstreamDrift_mm,
    rCenterAtCaptureX_mm => rUpstreamCenterX,
    rCenterAtCaptureY_mm => rUpstreamCenterY,
    rCenterNowX_mm => rUpstreamNowX,
    rCenterNowY_mm => rUpstreamNowY,
    rToRobotWorkStart_mm => rToRobotWorkStart_mm,
    aCornerNow => aUpstreamCornerNow
);
IF fbVisionResultEdge.Q THEN
    bExposureEncoderLatched := FALSE;
END_IF;
IF bUpstreamReset THEN
    bUpstreamReset := FALSE;
END_IF;

// ================================================================
// 8A. CAMERA PRODUCT FIFO — data only, no gantry motion commands.
// Real camera must provide CenterX/Y in millimeters, Angle in degrees.
// One unmatched exposure max (until camera provides explicit FrameID).
// Simulation requires bQueueSimMode and is isolated from QD75 Publisher.
// ================================================================
fbCameraQueue(
    bReset := bQueueReset OR bSystemStopRequested,
    bLiveExposure := bCameraExposeTrigger AND bSystemEStopOK,
    bLiveResult := bCameraTrigger AND bSystemEStopOK,
    bLiveBridgeVerified := bVisionFeedVerified,
    bCalibrationConfirmed := bVisionCalibrationOK,
    bSimMode := bQueueSimMode AND bSystemEStopOK AND NOT bLegacyMotionPublisherAllow
                AND NOT bXYManualPermit AND NOT bDebugXYPermit
                AND NOT bAutoDispatchEnable AND NOT bStartGlueCycle,
    bSimExposure := bQueueSimExposure AND bSystemEStopOK,
    bSimResult := bQueueSimResult AND bSystemEStopOK,
    bSimCompleteHead := bQueueSimCompleteHead AND bSystemEStopOK,
    rCenterX_mm := rCameraCenterX,
    rCenterY_mm := rCameraCenterY,
    rAngle_deg := rCameraAngleDeg,
    rCameraToWorkStart_mm := rCameraToWorkStart_mm,
    rCameraFineOffsetX_mm := rCamToRobotX_mm,
    rCameraOffsetY_mm := rCamToRobotY_mm,
    rCameraYaw_deg := rCamToRobotYaw_deg,
    rLength_mm := rProductLength,
    rWidth_mm := rProductWidth,
    rEncoderTotalDist_mm := rConveyorDist,
    rConveyorSpeed_mm_s := rConveyorSpeed,
    rXMin_mm := 0.0,
    rXMax_mm := 180.0,
    rYMin_mm := 0.0,
    rYMax_mm := 170.0,
    rMinCycleBudget_s := 1.2,
    rFlyTime_s := 0.12,
    rSyncTime_s := 0.06,
    nQueueCount => nQueueCount,
    nHeadProductID => nQueueHeadProductID,
    nHeadState => nQueueHeadState,
    bHeadValid => bQueueHeadValid,
    bHeadAllInside => bQueueHeadAllInside,
    bHeadForecastOK => bQueueHeadForecastOK,
    rHeadTravel_mm => rQueueHeadTravel_mm,
    rHeadToWorkStart_mm => rQueueToWorkStart_mm,
    rHeadCenterX_mm => rQueueHeadX_mm,
    rHeadCenterY_mm => rQueueHeadY_mm,
    aHeadCornerNow => aQueueHeadCornerNow,
    nAccepted => nQueueAccepted,
    nRejected => nQueueRejected,
    nMissed => nQueueMissed,
    nSimCompleted => nQueueSimCompleted,
    bInputFault => bQueueInputFault,
    nErrorCode => nQueueErrorCode
);

IF bQueueReset THEN
    bQueueReset := FALSE;
END_IF;

// ================================================================
// 9. DATA-ONLY PLC PUBLISH, wait for MANUAL ACK from audited spare M.
// Absolutely no robot Start/Move or M1001 spoofing from TwinCAT.
// ================================================================
bXYManualSafe := bSystemEStopOK AND NOT bDebugXYPermit
    AND NOT bGlueCycleBusy AND NOT bStartGlueCycle
    AND NOT bAbortGlueCycle AND NOT bGlueCycleError
    AND NOT bEnableManualWrite AND NOT bEchoPermit
    AND NOT bEchoWordBusy AND NOT bEchoBitBusy
    AND NOT bAutoDispatchEnable AND NOT bAutoDispatchArm
    AND NOT bTest_WriteM1000 AND NOT bTest_WriteD100
    AND (fbPublisher.nState = 0)
    AND bPlcQConnected;

fbXYManualAck(
    stSession := stMelsec,
    bExecute := bXYManualExecute AND bSystemEStopOK,
    bPermit := bXYManualPermit AND bSystemEStopOK AND bVisionFeedVerified
               AND bVisionCalibrationOK AND bXYManualSafe,
    bAckBitAudited := bXYManualAckBitAudited,
    nAckAddress := nXYManualAckMAddress,
    bSafeToWriteXY := bXYManualSafe,
    bProductCaptured := bUpstreamCaptured,
    aCornerNow := aUpstreamCornerNow,
    rConveyorSpeed := rConveyorSpeed,
    rFlyTime_s := 0.12,
    rXMax_mm := 180.0,
    rYMax_mm := 170.0,
    bAbort := bXYManualAbort OR bSystemStopRequested,
    bBusy => bXYManualBusy,
    bDone => bXYManualDone,
    bError => bXYManualError,
    nErrorCode => nXYManualErrorCode,
    nCommError => nXYManualCommError,
    nState => nXYManualState,
    nVertex => nXYManualVertex,
    nAckedVertices => nXYManualAcked,
    nSentX => nXYManualSentX,
    nSentY => nXYManualSentY,
    nReadX => nXYManualReadX,
    nReadY => nXYManualReadY,
    nReadVertex => nXYManualReadVertex,
    bReadbackOK => bXYManualReadbackOK,
    bRestored => bXYManualRestored
);

END_PROGRAM

// ---- POUs/FB_MelsecTcpConfig.TcPOU
FUNCTION_BLOCK FB_MelsecTcpConfig
VAR_INPUT
    bEnable         : BOOL := TRUE;                 // TRUE = duy trì kết nối
    sRemoteHost     : STRING(15) := '192.168.3.39'; // IP PLC-Q
    nRemotePort     : UDINT := 5010;               // Port MC Protocol
END_VAR
VAR_IN_OUT
    stSession       : ST_MelsecSession;             // Session TCP dùng chung
END_VAR
VAR
    fbConnect       : FB_SocketConnect;
    fbClose         : FB_SocketClose;
    tonRetry        : TON;

    nState          : INT := 0;
    bConnectError   : BOOL;
    nConnectErrorID : UDINT;
    bCloseError     : BOOL;
    nCloseErrorID   : UDINT;
    nReconnectCount : UDINT;
END_VAR

// State:
// 0 = chờ reconnect
// 1 = phát cạnh mở TCP
// 2 = chờ kết quả kết nối
// 10 = đã kết nối
// 20 = đóng socket khi Disable

CASE nState OF

    0: // Wait before reconnect. Never discard a live socket handle.
        stSession.bConnected := FALSE;

        IF NOT bEnable THEN
            tonRetry(IN := FALSE);
            stSession.bError := FALSE;
        ELSE
            // Backoff avoids an endless stream of new SYN requests when PLC has no slot.
            tonRetry(IN := TRUE, PT := T#5S);

            IF tonRetry.Q THEN
                tonRetry(IN := FALSE);
                stSession.bError := FALSE;
                nReconnectCount := nReconnectCount + 1;
                nState := 1;
            END_IF
        END_IF


    1: // Cạnh lên mở TCP Socket
        fbConnect(
            sSrvNetId   := '',
            sRemoteHost := sRemoteHost,
            nRemotePort := nRemotePort,
            bExecute    := TRUE,
            tTimeout    := T#35S,
            bError      => bConnectError,
            nErrId      => nConnectErrorID,
            hSocket     => stSession.hSocket
        );

        stSession.bBusy := TRUE;
        nState := 2;


    2: // Chờ FB_SocketConnect hoàn thành
        fbConnect(
            sSrvNetId   := '',
            sRemoteHost := sRemoteHost,
            nRemotePort := nRemotePort,
            bExecute    := FALSE,
            tTimeout    := T#35S,
            bError      => bConnectError,
            nErrId      => nConnectErrorID,
            hSocket     => stSession.hSocket
        );

        IF NOT fbConnect.bBusy THEN
            stSession.bBusy := FALSE;

            IF bConnectError THEN
                stSession.bError := TRUE;
                stSession.nErrorID := nConnectErrorID;
                stSession.bConnected := FALSE;
                // Do not zero a handle without trying to close it first.
                IF stSession.hSocket.handle <> 0 THEN
                    nState := 20;
                ELSE
                    nState := 0;
                END_IF;
            ELSE
                stSession.bConnected := TRUE;
                stSession.bError     := FALSE;
                stSession.nErrorID := 0;
                nState := 10;
            END_IF
        END_IF


    10: // Reconnect only after the read/write transaction releases the socket.
        IF NOT bEnable OR NOT stSession.bConnected THEN
            IF NOT stSession.bBusy THEN
                nState := 20;
            END_IF;
        END_IF


    20: // Close stale or disabled socket before any reconnect attempt.
        IF stSession.hSocket.handle = 0 THEN
            stSession.bConnected := FALSE;
            nState := 0;
        ELSE
            fbClose(
                sSrvNetId := '',
                hSocket := stSession.hSocket,
                bExecute := TRUE,
                tTimeout := T#5S,
                bError => bCloseError,
                nErrId => nCloseErrorID
            );
            nState := 21;
        END_IF;


    21: // Wait for close acknowledgement; keep an error for diagnostics.
        fbClose(
            sSrvNetId := '',
            hSocket := stSession.hSocket,
            bExecute := FALSE,
            tTimeout := T#5S,
            bError => bCloseError,
            nErrId => nCloseErrorID
        );

        IF NOT fbClose.bBusy THEN
            IF bCloseError THEN
                stSession.bError := TRUE;
                stSession.nErrorID := nCloseErrorID;
            END_IF;
            stSession.hSocket.handle := 0;
            stSession.bConnected := FALSE;
            nState := 0;
        END_IF

END_CASE

END_FUNCTION_BLOCK

// ---- POUs/FB_ConveyorEncoder.TcPOU
FUNCTION_BLOCK FB_ConveyorEncoder
VAR_INPUT
    bByte0          : BYTE;             // GVL.aIn[0]
    bByte1          : BYTE;             // GVL.aIn[1]
    rK_mm           : LREAL := 0.476475;// mm / xung (D=54.6mm, 360 xung)
    rCycleTime      : LREAL := 0.01;    // 10ms
END_VAR
VAR_OUTPUT
    nRawPulse       : UINT;             // Xung tức thời
    nDeltaPulse     : INT;              // Lệch xung mỗi 10ms
    rSpeed_mm_s     : LREAL;            // VẬN TỐC LỌC MƯỢT (mm/s)
    rSpeed_m_min    : LREAL;            // Vận tốc hiển thị (m/phút)
    rTotalDist_mm   : LREAL;            // TỔNG QUÃNG ĐƯỜNG (mm)
END_VAR
VAR
    nPrev           : UINT;
    bInit           : BOOL := TRUE;
    // 10 scan * 10ms = 100ms (theo interface contract)
    aDeltaBuf       : ARRAY[0..9] OF INT;
    nBufIdx         : INT := 0;
    nSumDelta       : DINT; // DINT để tránh tràn khi cộng nhiều xung
    nDelta32        : DINT;
END_VAR

// 1. Ghép 2 byte thành số xung 16-bit
nRawPulse := BYTE_TO_UINT(bByte1) * 256 + BYTE_TO_UINT(bByte0);

IF bInit THEN
    nPrev := nRawPulse;
    bInit := FALSE;
END_IF;

// Sai phân modulo 16-bit: encoder đếm 65535 -> 0 vẫn là +1 xung.
nDelta32 := UINT_TO_DINT(nRawPulse) - UINT_TO_DINT(nPrev);
IF nDelta32 > 32767 THEN
    nDelta32 := nDelta32 - 65536;
ELSIF nDelta32 < -32768 THEN
    nDelta32 := nDelta32 + 65536;
END_IF;
nDeltaPulse := DINT_TO_INT(nDelta32);
nPrev := nRawPulse;

// Rolling sum O(1), không quét cả bộ đệm trên mỗi scan.
nSumDelta := nSumDelta - INT_TO_DINT(aDeltaBuf[nBufIdx]) + nDelta32;
aDeltaBuf[nBufIdx] := nDeltaPulse;
nBufIdx := (nBufIdx + 1) MOD 10;

// Không làm tròn tốc độ sử dụng để tính tọa độ đón đầu.
IF rCycleTime > 0.0 THEN
    rSpeed_mm_s := DINT_TO_LREAL(nSumDelta) * rK_mm / (10.0 * rCycleTime);
ELSE
    rSpeed_mm_s := 0.0;
END_IF;
rSpeed_m_min := rSpeed_mm_s * 0.060;

rTotalDist_mm := rTotalDist_mm + DINT_TO_LREAL(nDelta32) * rK_mm;

END_FUNCTION_BLOCK

// ---- POUs/FB_InovanceMD200Conveyor.TcPOU
FUNCTION_BLOCK FB_InovanceMD200Conveyor
VAR_INPUT
    bEStopOK            : BOOL := FALSE; // NC safety chain feedback TRUE only when healthy
    bStart              : BOOL := FALSE; // operator START request, rising edge required
    rFrequencySet_Hz    : LREAL := 0.0;  // desired frequency, internally limited 0..25Hz
END_VAR
VAR_OUTPUT
    bDO_RunForward      : BOOL;          // ST-2318 Module 10 DO0 / pin 0
    nAO_12bitRaw        : INT;           // ST-4424 Module 11 AO1 12-bit 0..4095
    rAO_Volts           : LREAL;         // displayed expected 0..5V for 0..25Hz
    rTarget_Hz          : LREAL;
    rRamped_Hz          : LREAL;
    bAtTarget           : BOOL;
    bLimited25Hz        : BOOL;
    nStatus             : UINT;          // 0=STOP,1=RUN,2=ESTOP,3=RESTART_REQUIRED,4=BAD_FREQ
END_VAR
VAR
    fbStartRise         : R_TRIG;
    bFirstScan          : BOOL := TRUE;
    bStopSeen           : BOOL := FALSE;
    bRunGranted         : BOOL := FALSE;
    rStep               : LREAL;
    rDelta              : LREAL;
END_VAR
VAR CONSTANT
    cMaxFrequency_Hz    : LREAL := 25.0;  // fixed application limit
    cAnalogFullScale_Hz : LREAL := 50.0;  // verify MD200 0..10V => 0..50Hz
    cRampUp_HzPerS      : LREAL := 2.0;   // application reference ramp
    cTaskCycle_s        : LREAL := 0.01;  // must match PLC task period (10ms)
END_VAR

// Simplified MD200 controls: EStopOK + Start + Hz setpoint only.
// Safety-warning: EStopOK is an auxiliary status MONITOR, NOT a safety function.
// The machine's hardwired E-stop safety circuit must stop the drive independently.
// This FB is intentionally staged offline; do not Activate from a remote session.
//
// PLC boot, EStop loss or zero setpoint all revoke running authorization.
// Releasing EStop alone NEVER restarts a conveyor with START stuck TRUE.
// STOP must be observed and then START newly asserted.
fbStartRise(CLK := bStart);
IF bFirstScan THEN
    bFirstScan := FALSE;
    bStopSeen := FALSE;
    bRunGranted := FALSE;
    rRamped_Hz := 0.0;
END_IF;

// Outputs default safe every scan.
bDO_RunForward := FALSE;
nAO_12bitRaw := 0;
rAO_Volts := 0.0;
bAtTarget := FALSE;
bLimited25Hz := FALSE;
nStatus := 0;
rTarget_Hz := 0.0;

// Reject NaN: comparisons against NaN are invalid.
IF (rFrequencySet_Hz <> rFrequencySet_Hz) THEN
    bRunGranted := FALSE;
    rRamped_Hz := 0.0;
    nStatus := 4;
ELSE
    IF rFrequencySet_Hz > cMaxFrequency_Hz THEN
        rTarget_Hz := cMaxFrequency_Hz;
        bLimited25Hz := TRUE;
    ELSIF rFrequencySet_Hz > 0.0 THEN
        rTarget_Hz := rFrequencySet_Hz;
    ELSE
        rTarget_Hz := 0.0;
    END_IF;

    IF NOT bStart THEN
        bStopSeen := TRUE;
        bRunGranted := FALSE;
    END_IF;
    IF NOT bEStopOK OR (rTarget_Hz < 0.05) THEN
        bRunGranted := FALSE;
    END_IF;
    IF fbStartRise.Q AND bStopSeen AND bEStopOK AND (rTarget_Hz >= 0.05) THEN
        bRunGranted := TRUE;
    END_IF;

    IF NOT bEStopOK THEN
        nStatus := 2; // EStop healthy feedback missing
        rRamped_Hz := 0.0;
    ELSIF NOT bStart OR (rTarget_Hz < 0.05) THEN
        nStatus := 0;
        rRamped_Hz := 0.0;
    ELSIF NOT bRunGranted THEN
        nStatus := 3; // wait for STOP then fresh START edge
        rRamped_Hz := 0.0;
    ELSE
        nStatus := 1;
        rDelta := rTarget_Hz - rRamped_Hz;
        rStep := cRampUp_HzPerS * cTaskCycle_s;
        IF ABS(rDelta) <= rStep THEN
            rRamped_Hz := rTarget_Hz;
        ELSIF rDelta > 0.0 THEN
            rRamped_Hz := rRamped_Hz + rStep;
        ELSE
            rRamped_Hz := rRamped_Hz - rStep;
        END_IF;
        IF rRamped_Hz > cMaxFrequency_Hz THEN
            rRamped_Hz := cMaxFrequency_Hz;
        ELSIF rRamped_Hz < 0.0 THEN
            rRamped_Hz := 0.0;
        END_IF;
        rAO_Volts := (rRamped_Hz / cAnalogFullScale_Hz) * 10.0;
        nAO_12bitRaw := LREAL_TO_INT((rRamped_Hz / cAnalogFullScale_Hz) * 4095.0);
        IF nAO_12bitRaw > 4095 THEN nAO_12bitRaw := 4095; END_IF;
        IF nAO_12bitRaw < 0 THEN nAO_12bitRaw := 0; END_IF;
        bDO_RunForward := TRUE;
        bAtTarget := ABS(rTarget_Hz - rRamped_Hz) <= 0.0001;
    END_IF;
END_IF;

END_FUNCTION_BLOCK

// ---- POUs/FB_EziServoControl.TcPOU
FUNCTION_BLOCK FB_EziServoControl
VAR_INPUT
    bEnable         : BOOL := FALSE;
    bResetFault     : BOOL := FALSE;
    bJogFwd         : BOOL := FALSE;
    bJogBwd         : BOOL := FALSE;
    rTargetVelocity : LREAL := 100.0;
    rAcc            : LREAL := 400.0;
    rDec            : LREAL := 400.0;
END_VAR
VAR_IN_OUT
    Axis            : AXIS_REF;
END_VAR
VAR_OUTPUT
    bReady          : BOOL;
    rActPos_Deg     : LREAL;
    rActVel_Deg     : LREAL;
END_VAR
VAR
    fbPower         : MC_Power;
    fbMoveVelocity  : MC_MoveVelocity;
    fbHalt          : MC_Halt;
    fbReset         : MC_Reset;

    rTargetVel_Prev : LREAL;
    bVelChanged     : BOOL;
    fbTrigFwd       : R_TRIG;
    fbTrigBwd       : R_TRIG;
    fbTrigStop      : R_TRIG;
END_VAR

fbReset(Axis := Axis, Execute := bResetFault);

fbPower(
    Axis            := Axis,
    Enable          := bEnable,
    Enable_Positive := TRUE,
    Enable_Negative := TRUE,
    Override        := 100.0,
    Status          => bReady
);

fbTrigFwd(CLK := bEnable AND bJogFwd AND NOT bJogBwd);
fbTrigBwd(CLK := bEnable AND bJogBwd AND NOT bJogFwd);
fbTrigStop(CLK := NOT bEnable OR (NOT bJogFwd AND NOT bJogBwd) OR (bJogFwd AND bJogBwd));

IF rTargetVelocity <> rTargetVel_Prev THEN
    bVelChanged     := TRUE;
    rTargetVel_Prev := rTargetVelocity;
ELSE
    bVelChanged     := FALSE;
END_IF

fbMoveVelocity(
    Axis         := Axis,
    Execute      := (fbTrigFwd.Q OR fbTrigBwd.Q OR (bVelChanged AND (bJogFwd OR bJogBwd))),
    Velocity     := rTargetVelocity,
    Acceleration := rAcc,
    Deceleration := rDec,
    Jerk         := 10000.0,
    Direction    := SEL(bJogBwd, MC_Positive_Direction, MC_Negative_Direction)
);

fbHalt(
    Axis         := Axis,
    Execute      := fbTrigStop.Q,
    Deceleration := rDec,
    Jerk         := 10000.0
);

rActPos_Deg := Axis.NcToPlc.ActPos;
rActVel_Deg := Axis.NcToPlc.ActVelo;

END_FUNCTION_BLOCK

// ---- POUs/FB_ConveyorTracking4Pt.TcPOU
FUNCTION_BLOCK FB_ConveyorTracking4Pt
VAR_INPUT
    bResetSystem     : BOOL;
    bCameraResult    : BOOL;
    bAcceptCamera    : BOOL := TRUE;
    rCenterX_mm      : LREAL;
    rCenterY_mm      : LREAL;
    rAngleDeg        : LREAL;
    rLength_mm       : LREAL := 40.0;
    rWidth_mm        : LREAL := 40.0;
    nEncoderNow      : UINT;
    rMmPerPulse      : LREAL := 0.476475;
    rXMaxLimit_mm    : LREAL := 180.0;
END_VAR

VAR_OUTPUT
    bProductValid    : BOOL;
    nPulseAtCamera   : UINT;
    nPulseTravel     : INT;
    rTravel_mm       : LREAL;
    aCornerBase      : ARRAY[1..4] OF ST_Point2D;
    aCornerNow       : ARRAY[1..4] OF ST_Point2D;
END_VAR

VAR
    fbCameraEdge     : R_TRIG;
    rRad             : LREAL;
    rCosA            : LREAL;
    rSinA            : LREAL;
    rHalfLength      : LREAL;
    rHalfWidth       : LREAL;
    nIndex           : INT;
    bFirstScan       : BOOL := TRUE;
    nTravelRaw       : DINT;
END_VAR

// Reset mốc phần mềm một lần khi PLC khởi động hoặc khi bResetSystem kích.
IF bFirstScan OR bResetSystem THEN
    bFirstScan     := FALSE;
    bProductValid  := FALSE;
    nPulseAtCamera := nEncoderNow;
    nPulseTravel   := 0;
    rTravel_mm     := 0.0;

    FOR nIndex := 1 TO 4 DO
        aCornerBase[nIndex].X := 0.0;
        aCornerBase[nIndex].Y := 0.0;
        aCornerNow[nIndex].X  := 0.0;
        aCornerNow[nIndex].Y  := 0.0;
    END_FOR;
END_IF;

fbCameraEdge(CLK := bCameraResult);

// Camera chụp: chốt encoder và tính bốn góc gốc.
IF fbCameraEdge.Q AND bAcceptCamera THEN
    nPulseAtCamera := nEncoderNow;
    nPulseTravel   := 0;
    rTravel_mm     := 0.0;

    rRad   := rAngleDeg * 3.141592653589793 / 180.0;
    rCosA  := COS(rRad);
    rSinA  := SIN(rRad);
    rHalfLength := rLength_mm / 2.0;
    rHalfWidth  := rWidth_mm / 2.0;

    aCornerBase[1].X := rCenterX_mm + rHalfLength * rCosA - rHalfWidth * rSinA;
    aCornerBase[1].Y := rCenterY_mm + rHalfLength * rSinA + rHalfWidth * rCosA;
    aCornerBase[2].X := rCenterX_mm - rHalfLength * rCosA - rHalfWidth * rSinA;
    aCornerBase[2].Y := rCenterY_mm - rHalfLength * rSinA + rHalfWidth * rCosA;
    aCornerBase[3].X := rCenterX_mm - rHalfLength * rCosA + rHalfWidth * rSinA;
    aCornerBase[3].Y := rCenterY_mm - rHalfLength * rSinA - rHalfWidth * rCosA;
    aCornerBase[4].X := rCenterX_mm + rHalfLength * rCosA + rHalfWidth * rSinA;
    aCornerBase[4].Y := rCenterY_mm + rHalfLength * rSinA - rHalfWidth * rCosA;

    FOR nIndex := 1 TO 4 DO
        aCornerNow[nIndex] := aCornerBase[nIndex];
    END_FOR;
    bProductValid := TRUE;
END_IF;

// Tracking thời gian thực theo encoder.
IF bProductValid THEN
    nTravelRaw := UINT_TO_DINT(nEncoderNow) - UINT_TO_DINT(nPulseAtCamera);
    IF nTravelRaw > 32767 THEN
        nTravelRaw := nTravelRaw - 65536;
    ELSIF nTravelRaw < -32768 THEN
        nTravelRaw := nTravelRaw + 65536;
    END_IF;
    nPulseTravel := DINT_TO_INT(nTravelRaw);
    rTravel_mm   := TO_LREAL(nPulseTravel) * rMmPerPulse;

    FOR nIndex := 1 TO 4 DO
        aCornerNow[nIndex].X := aCornerBase[nIndex].X + rTravel_mm;
        aCornerNow[nIndex].Y := aCornerBase[nIndex].Y;
    END_FOR;

    // Hủy sản phẩm nếu toàn bộ cạnh phía sau đã vượt vùng X của Gantry.
    IF (aCornerNow[2].X > rXMaxLimit_mm) AND (aCornerNow[3].X > rXMaxLimit_mm) THEN
        bProductValid := FALSE;
        nPulseTravel  := 0;
        rTravel_mm    := 0.0;
    END_IF;
END_IF;

END_FUNCTION_BLOCK

// ---- POUs/FB_QD75CommandPublisher.TcPOU
FUNCTION_BLOCK FB_QD75CommandPublisher
VAR_INPUT
    // ================================================================
    // 1. ĐIỀU KHIỂN CHU TRÌNH TỰ ĐỘNG 4 ĐỈNH
    // ================================================================
    bStartCycle         : BOOL;             // Cạnh lên: bắt đầu chu trình 4 đỉnh
    bProductValid       : BOOL;            // Camera snapshot must exist before Start
    rEncoderDist_mm     : LREAL;           // Continuous conveyor distance from encoder
    bResetFault         : BOOL;            // Operator acknowledgement after fault
    bEnableManualWrite  : BOOL := FALSE;   // Deliberate service mode, OFF by default
    bAbortCycle         : BOOL;             // Hủy chu trình / yêu cầu dừng qua mạng

    // Dữ liệu từ khối Tracking & Băng tải
    aCornerNow          : ARRAY[1..4] OF ST_Point2D;
    rConveyorSpeed_mm_s : LREAL;

    // Thông số Gantry & Bù trôi
    rFlyTime_s          : LREAL := 0.120;  // Thời gian Gantry bay tiếp cận (120ms)
    rApproachSpeed_mm_s : LREAL := 500.0;  // Tốc độ bay tiếp cận (500 mm/s)
    rSyncTime_s         : LREAL := 0.060;  // Thời gian trượt đồng tốc X (60ms)
    rZDown_mm           : LREAL := 4.0;    // Độ cao Z hạ xuống chấm keo (4.0mm)
    rZSafe_mm           : LREAL := 0.0;    // Độ cao Z rút lên an toàn (0.0mm)

    // ================================================================
    // 2. CHẾ ĐỘ TEST THỦ CÔNG TRỰC TIẾP (KHI bStartCycle = FALSE)
    // ================================================================
    bManualWriteD100    : BOOL := FALSE;    // Click đúp TRUE -> Ghi số 32-bit vào D100-D101
    nD100_ManualVal     : DINT := 100;      // Giá trị 32-bit tùy ý bạn muốn ghi thử vào D100
    bManualWriteM1000   : BOOL := FALSE;    // Click đúp TRUE -> Ghi bit M1000 (ON hoặc OFF)
    bM1000_ManualVal    : BOOL := TRUE;     // TRUE = Bật M1000 ON, FALSE = Tắt M1000 OFF
    bManualReadM1001    : BOOL := FALSE;    // Click đúp TRUE -> Đọc bit M1001 từ PLC-Q về
END_VAR

VAR_IN_OUT
    stSession           : ST_MelsecSession; // Socket TCP dùng chung
END_VAR

VAR_OUTPUT
    // ================================================================
    // TRẠNG THÁI VÀ ĐẦU RA GIÁM SÁT
    // ================================================================
    stCommand           : ST_QD75_Command;  // Gói 15 words gửi sang D100..D114
    bCmdM1000           : BOOL;             // Trạng thái bit M1000
    bCmdM105            : BOOL;             // Trạng thái bit M105 (Abort)
    bBusy               : BOOL;             // Đang chạy chu trình 4 đỉnh
    bDone               : BOOL;             // Đã hoàn thành cả 4 đỉnh
    bError              : BOOL;             // Báo lỗi
    nErrorCode          : INT;              // Mã lỗi (501..503, 900..921)
    nCurrentVertex      : INT;              // Đỉnh đang thực hiện (1..4)

    rTargetX_mm         : LREAL;            // Tọa độ X đón đầu (mm)
    rTargetY_mm         : LREAL;            // Tọa độ Y (mm)
    rLead_mm            : LREAL;            // Bù trôi trong thời gian bay (mm)
    rDeltaXSync_mm      : LREAL;            // Quãng trượt đồng tốc X (mm)

    nLastCommError      : UDINT;            // MC socket/end-code diagnostics
    bM1001_ReadBack     : BOOL;             // Giá trị M1001 đọc được từ PLC-Q
    bStopCommandConfirmed : BOOL;           // Chỉ TRUE khi ghi M1000=OFF và M105=ON đều được ACK
END_VAR

VAR
    fbWrite             : FB_MelsecWrite;
    fbRead              : FB_MelsecRead;

    // Biến đệm dữ liệu truyền thông
    bM1000_Value        : BOOL;
    bM105_Value         : BOOL;
    bStatusBit          : BOOL;
    aStatusBits         : ARRAY[0..2] OF BOOL; // M102 Busy, M103 Position, M104 Alarm
    bM1000OffConfirmed  : BOOL;
    nD100_SendDINT      : DINT;

    // Tham số lệnh động
    bWriteReq           : BOOL;
    bReadReq            : BOOL;
    eWriteDevice        : E_MelsecDevice;
    nWriteAddress       : UDINT;
    nWritePoints        : UINT;
    bWriteBitMode       : BOOL;
    pWriteData          : PVOID;
    nWriteDataSize      : UDINT;

    eReadDevice         : E_MelsecDevice;
    nReadAddress        : UDINT;
    nReadPoints         : UINT;
    bReadBitMode        : BOOL;
    pReadData           : PVOID;
    nReadDataSize       : UDINT;

    nCommError          : UDINT;
    tonPoll             : TON;
    tonAck              : TON;            // Overall time limit, states 30+31
    tonRelease          : TON;            // Overall time limit, states 40+41
    aCycleCorners       : ARRAY[1..4] OF ST_Point2D;
    rCycleStartDist_mm  : LREAL;
    aRobotStatus        : ARRAY[0..2] OF BOOL; // M102 Busy, M103 InPosition, M104 Alarm
    tonStop             : TON;
    fbStartEdge         : R_TRIG;
    nState              : INT := 0;
END_VAR

fbStartEdge(CLK := bStartCycle);

// Update all watchdogs EVERY scan, including scans waiting for an asynchronous socket.
tonAck(IN := (nState = 30) OR (nState = 31) OR (nState = 33) OR (nState = 35), PT := T#10S);
tonRelease(IN := (nState = 40) OR (nState = 41) OR (nState = 43) OR (nState = 45), PT := T#5S);
tonStop(IN := (nState >= 90) AND (nState <= 92), PT := T#8S);

// Abort is a request through non-safety-rated TCP, NOT a hardware emergency stop.
IF bAbortCycle AND (nState <> 90) AND (nState <> 91)
    AND (nState <> 911) AND (nState <> 92)
    AND (nState <> 93) AND (nState <> 99) THEN
    bBusy := FALSE;
    bDone := FALSE;
    bError := TRUE;
    nErrorCode := 930;
    bStopCommandConfirmed := FALSE;
    nState := 90;
END_IF;

CASE nState OF
    0: // IDLE. No physical write occurs on transition to idle.
        bBusy := FALSE;
        bCmdM1000 := FALSE;
        nCurrentVertex := 0;
        bWriteReq := FALSE;
        bReadReq := FALSE;
        IF fbStartEdge.Q AND NOT bAbortCycle THEN
            IF NOT stSession.bConnected THEN
                bError := TRUE; nErrorCode := 900;
            ELSIF NOT bProductValid THEN
                bError := TRUE; nErrorCode := 901; // No valid camera product
            ELSIF stSession.bBusy THEN
                bError := TRUE; nErrorCode := 902; // Shared socket unavailable
            ELSE
                // Freeze identity of current product; use encoder travel for later vertices.
                aCycleCorners := aCornerNow;
                rCycleStartDist_mm := rEncoderDist_mm;
                bDone := FALSE; bError := FALSE; nErrorCode := 0;
                bBusy := TRUE; nCurrentVertex := 1;
                nState := 10;
            END_IF;
        ELSIF bManualWriteD100 OR bManualWriteM1000 THEN
            IF NOT bEnableManualWrite THEN
                bManualWriteD100 := FALSE;
                bManualWriteM1000 := FALSE;
                bError := TRUE; nErrorCode := 903; // Service mode disabled
            ELSIF stSession.bConnected AND NOT stSession.bBusy THEN
                IF bManualWriteD100 THEN
                    nD100_SendDINT := nD100_ManualVal;
                    eWriteDevice := DEV_D; nWriteAddress := 100; nWritePoints := 2;
                    bWriteBitMode := FALSE;
                    pWriteData := ADR(nD100_SendDINT); nWriteDataSize := SIZEOF(nD100_SendDINT);
                ELSE
                    bM1000_Value := bM1000_ManualVal;
                    eWriteDevice := DEV_M; nWriteAddress := 1000; nWritePoints := 1;
                    bWriteBitMode := TRUE;
                    pWriteData := ADR(bM1000_Value); nWriteDataSize := SIZEOF(bM1000_Value);
                END_IF;
                bWriteReq := TRUE; nState := 70;
            ELSE
                bManualWriteD100 := FALSE;
                bManualWriteM1000 := FALSE;
                bError := TRUE; nErrorCode := 900;
            END_IF;
        ELSIF bManualReadM1001 THEN
            IF stSession.bConnected AND NOT stSession.bBusy THEN
                eReadDevice := DEV_M; nReadAddress := 1001; nReadPoints := 1;
                bReadBitMode := TRUE;
                pReadData := ADR(bStatusBit); nReadDataSize := SIZEOF(bStatusBit);
                bReadReq := TRUE; nState := 80;
            ELSE
                bManualReadM1001 := FALSE;
                bError := TRUE; nErrorCode := 900;
            END_IF;
        END_IF;

    10: // Preflight before each vertex: read contiguous M102/M103/M104
        IF NOT stSession.bConnected THEN
            bError := TRUE; nErrorCode := 900; nState := 99;
        ELSE
            eReadDevice := DEV_M; nReadAddress := 102; nReadPoints := 3;
            bReadBitMode := TRUE;
            pReadData := ADR(aRobotStatus); nReadDataSize := SIZEOF(aRobotStatus);
            bReadReq := TRUE; nState := 11;
        END_IF;

    11:
        bReadReq := FALSE;
        IF fbRead.bDone THEN
            IF aRobotStatus[2] THEN
                bError := TRUE; nErrorCode := 904; nState := 99;
            ELSIF aRobotStatus[0] OR aRobotStatus[1] THEN
                bError := TRUE; nErrorCode := 905; nState := 99;
            ELSE
                nState := 14;
            END_IF;
        ELSIF fbRead.bError THEN
            nLastCommError := fbRead.nErrorID;
            bError := TRUE; nErrorCode := 920; nState := 99;
        END_IF;

    14: // ACK must also be low before any new command.
        eReadDevice := DEV_M; nReadAddress := 1001; nReadPoints := 1;
        bReadBitMode := TRUE;
        pReadData := ADR(bStatusBit); nReadDataSize := SIZEOF(bStatusBit);
        bReadReq := TRUE; nState := 15;

    15:
        bReadReq := FALSE;
        IF fbRead.bDone THEN
            IF bStatusBit THEN
                bError := TRUE; nErrorCode := 906; nState := 99;
            ELSE
                nState := 20;
            END_IF;
        ELSIF fbRead.bError THEN
            nLastCommError := fbRead.nErrorID;
            bError := TRUE; nErrorCode := 920; nState := 99;
        END_IF;

    20: // Validate every requested position BEFORE sending D100..D114.
        rLead_mm := rConveyorSpeed_mm_s * rFlyTime_s;
        rDeltaXSync_mm := rConveyorSpeed_mm_s * rSyncTime_s;
        rTargetX_mm := aCycleCorners[nCurrentVertex].X
                       + (rEncoderDist_mm - rCycleStartDist_mm) + rLead_mm;
        rTargetY_mm := aCycleCorners[nCurrentVertex].Y;

        IF (nCurrentVertex < 1) OR (nCurrentVertex > 4)
            OR (rConveyorSpeed_mm_s <= 0.0) OR (rConveyorSpeed_mm_s > 1000.0)
            OR (rApproachSpeed_mm_s <= 0.0) OR (rApproachSpeed_mm_s > 1000.0)
            OR (rFlyTime_s < 0.0) OR (rFlyTime_s > 1.0)
            OR (rSyncTime_s <= 0.0) OR (rSyncTime_s > 0.5)
            OR (rTargetX_mm < 0.0) OR ((rTargetX_mm + rDeltaXSync_mm) > 180.0)
            OR (rTargetY_mm < 0.0) OR (rTargetY_mm > 170.0)
            OR (rZSafe_mm < 0.0) OR (rZDown_mm > 52.0)
            OR (rZDown_mm < rZSafe_mm) THEN
            bError := TRUE; nErrorCode := 501; nState := 99;
        ELSE
            stCommand.Target_X       := LREAL_TO_DINT(rTargetX_mm * 10000.0);
            stCommand.Target_Y       := LREAL_TO_DINT(rTargetY_mm * 10000.0);
            stCommand.Target_Z_Down  := LREAL_TO_DINT(rZDown_mm * 10000.0);
            stCommand.Target_Z_Safe  := LREAL_TO_DINT(rZSafe_mm * 10000.0);
            stCommand.Speed_Approach := LREAL_TO_DINT(rApproachSpeed_mm_s * 6000.0);
            stCommand.Speed_Sync     := LREAL_TO_DINT(rConveyorSpeed_mm_s * 6000.0);
            stCommand.DeltaX_Sync    := LREAL_TO_DINT(rDeltaXSync_mm * 10000.0);
            stCommand.Vertex_Index  := nCurrentVertex;

            eWriteDevice := DEV_D; nWriteAddress := 100; nWritePoints := 15;
            bWriteBitMode := FALSE;
            pWriteData := ADR(stCommand); nWriteDataSize := SIZEOF(stCommand);
            bWriteReq := TRUE; nState := 21;
        END_IF;

    21:
        bWriteReq := FALSE;
        IF fbWrite.bDone THEN
            // Tạo ít nhất một scan bExecute=FALSE trước lệnh ghi tiếp theo.
            nState := 211;
        ELSIF fbWrite.bError THEN
            nLastCommError := fbWrite.nErrorID;
            bError := TRUE; nErrorCode := 910; nState := 90;
        END_IF;

    211:
        bCmdM1000 := TRUE; bM1000_Value := TRUE;
        eWriteDevice := DEV_M; nWriteAddress := 1000; nWritePoints := 1;
        bWriteBitMode := TRUE;
        pWriteData := ADR(bM1000_Value); nWriteDataSize := SIZEOF(bM1000_Value);
        bWriteReq := TRUE; nState := 22;

    22:
        bWriteReq := FALSE;
        IF fbWrite.bDone THEN
            nState := 30;
        ELSIF fbWrite.bError THEN
            nLastCommError := fbWrite.nErrorID;
            bError := TRUE; nErrorCode := 911; nState := 90;
        END_IF;

    30:
        IF tonAck.Q THEN
            bError := TRUE; nErrorCode := 920; nState := 90;
        ELSE
            tonPoll(IN := TRUE, PT := T#20MS);
            IF tonPoll.Q THEN
                tonPoll(IN := FALSE);
                eReadDevice := DEV_M; nReadAddress := 104; nReadPoints := 1;
                bReadBitMode := TRUE;
                pReadData := ADR(aRobotStatus[2]); nReadDataSize := SIZEOF(aRobotStatus[2]);
                bReadReq := TRUE; nState := 33;
            END_IF;
        END_IF;

    33: // Giám sát M104 Alarm cả trong lúc chờ hoàn thành đỉnh.
        bReadReq := FALSE;
        IF fbRead.bDone THEN
            IF aRobotStatus[2] THEN
                bError := TRUE; nErrorCode := 927; nState := 90;
            ELSE
                nState := 35;
            END_IF;
        ELSIF fbRead.bError THEN
            bError := TRUE; nErrorCode := 928; nState := 90;
        END_IF;

    35:
        eReadDevice := DEV_M; nReadAddress := 1001; nReadPoints := 1;
        bReadBitMode := TRUE;
        pReadData := ADR(bStatusBit); nReadDataSize := SIZEOF(bStatusBit);
        bReadReq := TRUE; nState := 31;

    31:
        bReadReq := FALSE;
        IF tonAck.Q THEN
            bError := TRUE; nErrorCode := 920; nState := 90;
        ELSIF fbRead.bDone THEN
            bM1001_ReadBack := bStatusBit;
            IF bStatusBit THEN
                bCmdM1000 := FALSE; bM1000_Value := FALSE;
                eWriteDevice := DEV_M; nWriteAddress := 1000; nWritePoints := 1;
                bWriteBitMode := TRUE;
                pWriteData := ADR(bM1000_Value); nWriteDataSize := SIZEOF(bM1000_Value);
                bWriteReq := TRUE; nState := 32;
            ELSE
                nState := 30;
            END_IF;
        ELSIF fbRead.bError THEN
            nLastCommError := fbRead.nErrorID;
            bError := TRUE; nErrorCode := 920; nState := 90;
        END_IF;

    32:
        bWriteReq := FALSE;
        IF fbWrite.bDone THEN
            nState := 40;
        ELSIF fbWrite.bError THEN
            nLastCommError := fbWrite.nErrorID;
            bError := TRUE; nErrorCode := 912; nState := 90;
        END_IF;

    40:
        IF tonRelease.Q THEN
            bError := TRUE; nErrorCode := 921; nState := 90;
        ELSE
            tonPoll(IN := TRUE, PT := T#20MS);
            IF tonPoll.Q THEN
                tonPoll(IN := FALSE);
                eReadDevice := DEV_M; nReadAddress := 104; nReadPoints := 1;
                bReadBitMode := TRUE;
                pReadData := ADR(aRobotStatus[2]); nReadDataSize := SIZEOF(aRobotStatus[2]);
                bReadReq := TRUE; nState := 43;
            END_IF;
        END_IF;

    43:
        bReadReq := FALSE;
        IF fbRead.bDone THEN
            IF aRobotStatus[2] THEN
                bError := TRUE; nErrorCode := 927; nState := 90;
            ELSE
                nState := 45;
            END_IF;
        ELSIF fbRead.bError THEN
            bError := TRUE; nErrorCode := 928; nState := 90;
        END_IF;

    45:
        eReadDevice := DEV_M; nReadAddress := 1001; nReadPoints := 1;
        bReadBitMode := TRUE;
        pReadData := ADR(bStatusBit); nReadDataSize := SIZEOF(bStatusBit);
        bReadReq := TRUE; nState := 41;

    41:
        bReadReq := FALSE;
        IF tonRelease.Q THEN
            bError := TRUE; nErrorCode := 921; nState := 90;
        ELSIF fbRead.bDone THEN
            bM1001_ReadBack := bStatusBit;
            IF NOT bStatusBit THEN
                IF nCurrentVertex < 4 THEN
                    nCurrentVertex := nCurrentVertex + 1;
                    nState := 10; // Preflight next vertex, including M103 and M104
                ELSE
                    bBusy := FALSE; bDone := TRUE; nState := 0;
                END_IF;
            ELSE
                nState := 40;
            END_IF;
        ELSIF fbRead.bError THEN
            nLastCommError := fbRead.nErrorID;
            bError := TRUE; nErrorCode := 921; nState := 90;
        END_IF;

    70: // Manual write (service mode only)
        bWriteReq := FALSE;
        IF fbWrite.bDone OR fbWrite.bError THEN
            IF fbWrite.bError THEN
                nLastCommError := fbWrite.nErrorID;
                bError := TRUE; nErrorCode := 910;
            END_IF;
            bManualWriteD100 := FALSE; bManualWriteM1000 := FALSE;
            nState := 0;
        END_IF;

    80: // Read-only diagnostics
        bReadReq := FALSE;
        IF fbRead.bDone OR fbRead.bError THEN
            IF fbRead.bDone THEN
                bM1001_ReadBack := bStatusBit;
            ELSE
                nLastCommError := fbRead.nErrorID;
                bError := TRUE; nErrorCode := 920;
            END_IF;
            bManualReadM1001 := FALSE; nState := 0;
        END_IF;

    90: // Best-effort abort: wait for a pending transaction to finish first.
        bWriteReq := FALSE;
        bReadReq := FALSE;
        bBusy := FALSE; bDone := FALSE; bCmdM1000 := FALSE; bCmdM105 := TRUE;
        IF NOT stSession.bConnected OR tonStop.Q THEN
            bError := TRUE; nState := 99;
        ELSIF NOT stSession.bBusy AND NOT fbWrite.bBusy AND NOT fbRead.bBusy THEN
            bM105_Value := TRUE;
            eWriteDevice := DEV_M; nWriteAddress := 105; nWritePoints := 1;
            bWriteBitMode := TRUE;
            pWriteData := ADR(bM105_Value); nWriteDataSize := SIZEOF(bM105_Value);
            bWriteReq := TRUE; nState := 91;
        END_IF;

    91:
        bWriteReq := FALSE;
        IF fbWrite.bDone THEN
            nState := 911; // Ngắt một scan bExecute để R_TRIG ghi tiếp nhận cạnh lên.
        ELSIF fbWrite.bError OR tonStop.Q THEN
            nLastCommError := fbWrite.nErrorID;
            bError := TRUE; nState := 99;
        END_IF;

    911:
        bM1000_Value := FALSE;
        eWriteDevice := DEV_M; nWriteAddress := 1000; nWritePoints := 1;
        bWriteBitMode := TRUE;
        pWriteData := ADR(bM1000_Value); nWriteDataSize := SIZEOF(bM1000_Value);
        bWriteReq := TRUE; nState := 92;

    92:
        bWriteReq := FALSE;
        IF fbWrite.bDone THEN
            bStopCommandConfirmed := TRUE;
            bError := TRUE; nState := 99;
        ELSIF fbWrite.bError OR tonStop.Q THEN
            nLastCommError := fbWrite.nErrorID;
            bError := TRUE; nState := 99;
        END_IF;

    99: // Fault latched. No automatic restart, manual acknowledgement required.
        bBusy := FALSE;
        bWriteReq := FALSE;
        bReadReq := FALSE;
        IF bResetFault AND NOT bAbortCycle AND NOT bStartCycle AND stSession.bConnected
            AND NOT stSession.bBusy AND NOT fbWrite.bBusy AND NOT fbRead.bBusy THEN
            IF NOT bStopCommandConfirmed THEN
                nState := 90; // Chưa nhận ACK dừng: bắt buộc thử dừng lại trước khi reset.
            ELSE
            bM105_Value := FALSE; // Deliberate operator reset after safe conditions
            eWriteDevice := DEV_M; nWriteAddress := 105; nWritePoints := 1;
            bWriteBitMode := TRUE;
            pWriteData := ADR(bM105_Value); nWriteDataSize := SIZEOF(bM105_Value);
            bWriteReq := TRUE; nState := 95;
            END_IF;
        END_IF;

    95:
        bWriteReq := FALSE;
        IF fbWrite.bDone THEN
            bCmdM105 := FALSE; bCmdM1000 := FALSE;
            bStopCommandConfirmed := FALSE;
            bError := FALSE; nErrorCode := 0; nState := 0;
        ELSIF fbWrite.bError THEN
            nLastCommError := fbWrite.nErrorID;
            nState := 99;
        END_IF;
END_CASE;

// Exactly one operation at a time; both FBs use ownership-based socket locking.
fbWrite(
    stSession := stSession, bExecute := bWriteReq,
    eDevice := eWriteDevice, nStartAddr := nWriteAddress,
    nPoints := nWritePoints, bBitAccess := bWriteBitMode,
    pData := pWriteData, nDataSize := nWriteDataSize,
    nErrorID => nCommError
);
fbRead(
    stSession := stSession, bExecute := bReadReq,
    eDevice := eReadDevice, nStartAddr := nReadAddress,
    nPoints := nReadPoints, bBitAccess := bReadBitMode,
    pData := pReadData, nDataSize := nReadDataSize,
    nErrorID => nCommError
);

END_FUNCTION_BLOCK

// ---- POUs/FB_MelsecWrite.TcPOU
FUNCTION_BLOCK FB_MelsecWrite
VAR_INPUT
    bExecute    : BOOL;             // Cạnh lên: Bắt đầu giao dịch Write
    eDevice     : E_MelsecDevice;   // Mã vùng nhớ (DEV_D, DEV_M, ...)
    nStartAddr  : UDINT;            // Địa chỉ bắt đầu (D100 -> 100, M1000 -> 1000)
    nPoints     : UINT;             // Số điểm ghi (Số word hoặc số bit)
    bBitAccess  : BOOL;             // TRUE: Ghi bit (M), FALSE: Ghi word (D)
    pData       : PVOID;            // Con trỏ tới vùng dữ liệu nguồn
    nDataSize   : UDINT;            // Kích thước dữ liệu nguồn (bytes)
END_VAR

VAR_IN_OUT
    stSession   : ST_MelsecSession; // Session TCP dùng chung
END_VAR

VAR_OUTPUT
    bBusy       : BOOL;
    bDone       : BOOL;
    bError      : BOOL;
    nErrorID    : UDINT;            // 0=OK, Mã lỗi Beckhoff socket hoặc EndCode Mitsubishi
END_VAR

VAR
    fbTrigger   : R_TRIG;
    fbSend      : FB_SocketSend;
    fbReceive   : FB_SocketReceive;
    tonTimeout  : TON;

    aTx         : ARRAY[0..255] OF BYTE;
    aRx         : ARRAY[0..63] OF BYTE;
    nSendLength : UDINT;
    nWriteBytes : UDINT;
    nEndCode    : UINT;

    pSrcByte    : POINTER TO BYTE;
    pSrcBit     : POINTER TO BOOL;
    nIdx        : UDINT;
    nPairIdx    : UDINT;
    bBitVal1    : BYTE;
    bBitVal2    : BYTE;

    nRequestLength : UINT;
    nState      : INT := 0;
    bOwnsSession : BOOL;
    nRxCount    : UDINT;
    nExpectedFrame : UDINT;
END_VAR

fbTrigger(CLK := bExecute);
// Timer receives a scan on every PLC cycle, even between TCP polls.
tonTimeout(IN := bBusy AND ((nState = 20) OR (nState = 21)), PT := T#5S);

// Xóa cờ trạng thái khi bắt đầu lệnh mới
IF nState = 0 THEN
    IF fbTrigger.Q THEN
        bDone    := FALSE;
        bError   := FALSE;
        nErrorID := 0;
    END_IF;
END_IF;

// Kiểm tra điều kiện tiên quyết
IF fbTrigger.Q THEN
    IF NOT stSession.bConnected THEN
        bError   := TRUE;
        nErrorID := 16#E001; // Socket chưa kết nối
        RETURN;
    ELSIF stSession.bBusy THEN
        bError   := TRUE;
        nErrorID := 16#E002; // Kênh truyền đang bận
        RETURN;
    ELSIF (pData = 0) OR (nDataSize = 0) THEN
        bError   := TRUE;
        nErrorID := 16#E003; // Con trỏ dữ liệu không hợp lệ
        RETURN;
    ELSIF (nPoints = 0) OR (nStartAddr > 16#FFFFFF)
        OR (bBitAccess AND ((UINT_TO_UDINT(nPoints) > nDataSize) OR (((UINT_TO_UDINT(nPoints) + 1) / 2) > (SIZEOF(aTx) - 21))))
        OR ((NOT bBitAccess) AND (((UINT_TO_UDINT(nPoints) * 2) > nDataSize) OR ((UINT_TO_UDINT(nPoints) * 2) > (SIZEOF(aTx) - 21)))) THEN
        bError := TRUE;
        nErrorID := 16#E004; // Invalid quantity, address or source length
        RETURN;
    ELSE
        // ============================================================
        // 1. ĐÓNG GÓI KHUNG TRUYỀN MC PROTOCOL 3E FRAME (BINARY WRITE)
        // ============================================================
        // 1.1. Subheader: 0x50 0x00 (Gửi yêu cầu không giám sát)
        aTx[0] := 16#50;
        aTx[1] := 16#00;

        // 1.2. Network No: 0x00 (Mạng cục bộ)
        aTx[2] := 16#00;

        // 1.3. PC No: 0xFF (Trạm đích trực tiếp)
        aTx[3] := 16#FF;

        // 1.4. Target Module I/O No: 0xFF 0x03 (CPU đa xử lý mặc định)
        aTx[4] := 16#FF;
        aTx[5] := 16#03;

        // 1.5. Target Module Multidrop Station No: 0x00
        aTx[6] := 16#00;

        // Bytes 7..8: Request Data Length (sẽ tính và ghi sau khi nạp payload)

        // 1.6. Monitoring Timer: 0x10 0x00 (Đơn vị 250ms -> 16 = 4 giây)
        aTx[9]  := 16#10;
        aTx[10] := 16#00;

        // 1.7. Command: 0x01 0x14 (Batch Write - Ghi hàng loạt)
        aTx[11] := 16#01;
        aTx[12] := 16#14;

        // 1.8. Subcommand: 0x0001 (Bit units) hoặc 0x0000 (Word units)
        IF bBitAccess THEN
            aTx[13] := 16#01;
            aTx[14] := 16#00;
        ELSE
            aTx[13] := 16#00;
            aTx[14] := 16#00;
        END_IF;

        // 1.9. Start Device Address (3 bytes: LSB -> MSB)
        aTx[15] := UDINT_TO_BYTE(nStartAddr AND 16#FF);
        aTx[16] := UDINT_TO_BYTE(SHR(nStartAddr, 8) AND 16#FF);
        aTx[17] := UDINT_TO_BYTE(SHR(nStartAddr, 16) AND 16#FF);

        // 1.10. Device Code (M=0x90, D=0xA8, ...)
        aTx[18] := TO_BYTE(eDevice);

        // 1.11. Number of Device Points (2 bytes: LSB -> MSB)
        aTx[19] := UINT_TO_BYTE(nPoints AND 16#FF);
        aTx[20] := UINT_TO_BYTE(SHR(nPoints, 8) AND 16#FF);

        // ============================================================
        // 1.12. NẠP DỮ LIỆU CẦN GHI (WRITE PAYLOAD)
        // ============================================================
        IF bBitAccess THEN
            // Ghi Bit: MC Protocol mã hóa 2 bit vào 1 byte (Mỗi nibble 4-bit chứa 1 bit dữ liệu 0x10 / 0x01)
            pSrcBit := pData;
            nWriteBytes := (nPoints + 1) / 2; // Số byte payload

            FOR nPairIdx := 0 TO (nWriteBytes - 1) DO
                // Bit thứ nhất (nibble cao)
                IF (nPairIdx * 2) < nPoints THEN
                    IF pSrcBit[nPairIdx * 2] THEN
                        bBitVal1 := 16#10;
                    ELSE
                        bBitVal1 := 16#00;
                    END_IF;
                ELSE
                    bBitVal1 := 16#00;
                END_IF;

                // Bit thứ hai (nibble thấp)
                IF (nPairIdx * 2 + 1) < nPoints THEN
                    IF pSrcBit[nPairIdx * 2 + 1] THEN
                        bBitVal2 := 16#01;
                    ELSE
                        bBitVal2 := 16#00;
                    END_IF;
                ELSE
                    bBitVal2 := 16#00;
                END_IF;

                aTx[21 + nPairIdx] := bBitVal1 OR bBitVal2;
            END_FOR;

        ELSE
            // Ghi Word: Sao chép trực tiếp mảng bytes (Mỗi word = 2 bytes)
            pSrcByte := pData;
            nWriteBytes := UINT_TO_UDINT(nPoints) * 2;

            FOR nIdx := 0 TO (nWriteBytes - 1) DO
                aTx[21 + nIdx] := pSrcByte[nIdx];
            END_FOR;
        END_IF;

        // 1.13. Tính Request Data Length (Từ Monitoring Timer tới hết Payload)
        // Timer(2) + Cmd(2) + Subcmd(2) + Addr(3) + Dev(1) + Points(2) + Payload = 12 + nWriteBytes
        nRequestLength := 12 + UDINT_TO_UINT(nWriteBytes);
        aTx[7] := UINT_TO_BYTE(nRequestLength AND 16#FF);
        aTx[8] := UINT_TO_BYTE(SHR(nRequestLength, 8) AND 16#FF);

        // Tổng chiều dài khung gửi đi: Subheader(2) + Net(1) + PC(1) + IO(2) + Drop(1) + Len(2) + RequestLength
        nSendLength := 9 + nRequestLength;

        bBusy  := TRUE;
        bOwnsSession := TRUE;
        nRxCount := 0;
        nExpectedFrame := 0;
        nState := 10;
    END_IF;
END_IF;


// ================================================================
// MÁY TRẠNG THÁI GIAO TIẾP SOCKET
// ================================================================
CASE nState OF

    10: // Phát lệnh gửi dữ liệu qua TCP
        fbSend(
            sSrvNetId := '',
            hSocket   := stSession.hSocket,
            cbLen     := nSendLength,
            pSrc      := ADR(aTx),
            bExecute  := TRUE,
            tTimeout  := T#3S
        );

        nState := 11;


    11: // Chờ gửi xong
        fbSend(
            sSrvNetId := '',
            hSocket   := stSession.hSocket,
            cbLen     := nSendLength,
            pSrc      := ADR(aTx),
            bExecute  := FALSE,
            tTimeout  := T#3S
        );

        IF NOT fbSend.bBusy THEN
            IF fbSend.bError THEN
                bError   := TRUE;
                nErrorID := fbSend.nErrId;
                stSession.bConnected := FALSE;
                bBusy    := FALSE;
                nState   := 0;
            ELSE
                nState := 20;
            END_IF;
        END_IF;


    20: // Phát lệnh nhận phản hồi PLC
        fbReceive(
            sSrvNetId := '',
            hSocket   := stSession.hSocket,
            cbLen     := SIZEOF(aRx) - nRxCount,
            pDest     := ADR(aRx[nRxCount]),
            bExecute  := TRUE,
            tTimeout  := T#3S
        );

        nState := 21;


    21: // Chờ nhận phản hồi (Polled receive với timeout 2 giây)
        fbReceive(
            sSrvNetId := '',
            hSocket   := stSession.hSocket,
            cbLen     := SIZEOF(aRx) - nRxCount,
            pDest     := ADR(aRx[nRxCount]),
            bExecute  := FALSE,
            tTimeout  := T#3S
        );

        IF NOT fbReceive.bBusy THEN
            IF fbReceive.bError THEN
                bError   := TRUE;
                nErrorID := fbReceive.nErrId;
                stSession.bConnected := FALSE;
                bBusy    := FALSE;
                nState   := 0;

            ELSIF fbReceive.nRecBytes > 0 THEN
                nRxCount := nRxCount + fbReceive.nRecBytes;
                IF nRxCount >= 9 THEN
                    nExpectedFrame := 9 + BYTE_TO_UDINT(aRx[7]) + BYTE_TO_UDINT(aRx[8]) * 256;
                    IF (nExpectedFrame < 11) OR (nExpectedFrame > SIZEOF(aRx)) THEN
                        bError := TRUE; nErrorID := 16#E006;
                        stSession.bConnected := FALSE;
                        bBusy := FALSE; nState := 0;
                    ELSIF nRxCount >= nExpectedFrame THEN
                        IF (aRx[0] <> 16#D0) OR (aRx[1] <> 16#00) THEN
                            bError := TRUE; nErrorID := 16#E007;
                            stSession.bConnected := FALSE;
                        ELSE
                            nEndCode := BYTE_TO_UINT(aRx[9]) + BYTE_TO_UINT(aRx[10]) * 256;
                            IF nEndCode = 0 THEN
                                bDone := TRUE;
                            ELSE
                                bError := TRUE; nErrorID := nEndCode;
                            END_IF;
                        END_IF;
                        bBusy := FALSE; nState := 0;
                    ELSE
                        nState := 20; // Continue receiving fragmented response
                    END_IF;
                ELSE
                    nState := 20; // Header not yet complete
                END_IF;

            ELSIF tonTimeout.Q THEN
                // Quá 2 giây không có phản hồi
                bError   := TRUE;
                nErrorID := 16#E008; // Timeout chờ response PLC
                stSession.bConnected := FALSE;
                bBusy    := FALSE;
                nState   := 0;

            ELSE
                // Chưa có dữ liệu về trong scan này -> Kích đọc tiếp ở scan sau
                nState := 20;
            END_IF;
        END_IF;

END_CASE;

// Cập nhật trạng thái bận vào session dùng chung
// Only the FB that acquired the socket lock may release it.
IF bBusy THEN
    stSession.bBusy := TRUE;
ELSIF bOwnsSession THEN
    stSession.bBusy := FALSE;
    bOwnsSession := FALSE;
END_IF;

END_FUNCTION_BLOCK

// ---- POUs/FB_MelsecRead.TcPOU
FUNCTION_BLOCK FB_MelsecRead
VAR_INPUT
    bExecute    : BOOL;             // Cạnh lên: Bắt đầu giao dịch Read
    eDevice     : E_MelsecDevice;   // Loại vùng nhớ (DEV_M, DEV_D, ...)
    nStartAddr  : UDINT;            // Địa chỉ bắt đầu (M1001 -> 1001, D100 -> 100)
    nPoints     : UINT;             // Số điểm đọc (Số bit hoặc số word)
    bBitAccess  : BOOL;             // TRUE: Đọc Bit (M), FALSE: Đọc Word (D)
    pData       : PVOID;            // Con trỏ tới vùng đệm lưu kết quả đọc
    nDataSize   : UDINT;            // Kích thước vùng đệm đích (bytes)
END_VAR

VAR_IN_OUT
    stSession   : ST_MelsecSession; // Session TCP dùng chung
END_VAR

VAR_OUTPUT
    bBusy       : BOOL;
    bDone       : BOOL;
    bError      : BOOL;
    nErrorID    : UDINT;            // 0=OK, Mã lỗi Beckhoff socket hoặc EndCode Mitsubishi
END_VAR

VAR
    fbTrigger   : R_TRIG;
    fbSend      : FB_SocketSend;
    fbReceive   : FB_SocketReceive;
    tonTimeout  : TON;

    aTx         : ARRAY[0..31] OF BYTE;
    aRx         : ARRAY[0..255] OF BYTE;
    nEndCode    : UINT;

    pDestByte   : POINTER TO BYTE;
    pDestBit    : POINTER TO BOOL;
    nIdx        : UDINT;
    nCopyBytes  : UDINT;

    nState      : INT := 0;
    bOwnsSession : BOOL;
    nRxCount    : UDINT;
    nExpectedFrame : UDINT;
END_VAR

fbTrigger(CLK := bExecute);
// Timer receives a scan on every PLC cycle, even between TCP polls.
tonTimeout(IN := bBusy AND ((nState = 20) OR (nState = 21)), PT := T#5S);

// Xóa cờ trạng thái khi bắt đầu lệnh mới
IF nState = 0 THEN
    IF fbTrigger.Q THEN
        bDone    := FALSE;
        bError   := FALSE;
        nErrorID := 0;
    END_IF;
END_IF;

// Kiểm tra điều kiện tiên quyết
IF fbTrigger.Q THEN
    IF NOT stSession.bConnected THEN
        bError   := TRUE;
        nErrorID := 16#E101; // Socket chưa kết nối
        RETURN;
    ELSIF stSession.bBusy THEN
        bError   := TRUE;
        nErrorID := 16#E102; // Session đang bận
        RETURN;
    ELSIF (pData = 0) OR (nDataSize = 0) THEN
        bError   := TRUE;
        nErrorID := 16#E103; // Vùng đệm đích không hợp lệ
        RETURN;
    ELSIF (nPoints = 0) OR (nStartAddr > 16#FFFFFF)
        OR (bBitAccess AND ((UINT_TO_UDINT(nPoints) > nDataSize) OR (((UINT_TO_UDINT(nPoints) + 1) / 2) > (SIZEOF(aRx) - 11))))
        OR ((NOT bBitAccess) AND (((UINT_TO_UDINT(nPoints) * 2) > nDataSize) OR ((UINT_TO_UDINT(nPoints) * 2) > (SIZEOF(aRx) - 11)))) THEN
        bError := TRUE;
        nErrorID := 16#E106; // Invalid quantity, address or destination length
        RETURN;
    ELSE
        // ============================================================
        // 1. ĐÓNG GÓI KHUNG YÊU CẦU ĐỌC MC PROTOCOL 3E (BINARY READ)
        // Chiều dài cố định: 21 bytes
        // ============================================================
        // 1.1. Subheader: 0x50 0x00
        aTx[0] := 16#50;
        aTx[1] := 16#00;

        // 1.2. Network No: 0x00
        aTx[2] := 16#00;

        // 1.3. PC No: 0xFF
        aTx[3] := 16#FF;

        // 1.4. Target Module I/O: 0xFF 0x03
        aTx[4] := 16#FF;
        aTx[5] := 16#03;

        // 1.5. Target Module Drop: 0x00
        aTx[6] := 16#00;

        // 1.6. Request Data Length: 12 bytes (Từ Timer đến hết Points: 2+2+2+3+1+2 = 12)
        aTx[7] := 16#0C;
        aTx[8] := 16#00;

        // 1.7. Monitoring Timer: 0x10 0x00 (4 giây)
        aTx[9]  := 16#10;
        aTx[10] := 16#00;

        // 1.8. Command: 0x01 0x04 (Batch Read - Đọc hàng loạt)
        aTx[11] := 16#01;
        aTx[12] := 16#04;

        // 1.9. Subcommand: 0x0001 (Bit units) hoặc 0x0000 (Word units)
        IF bBitAccess THEN
            aTx[13] := 16#01;
            aTx[14] := 16#00;
        ELSE
            aTx[13] := 16#00;
            aTx[14] := 16#00;
        END_IF;

        // 1.10. Start Device Address (3 bytes: LSB -> MSB)
        aTx[15] := UDINT_TO_BYTE(nStartAddr AND 16#FF);
        aTx[16] := UDINT_TO_BYTE(SHR(nStartAddr, 8) AND 16#FF);
        aTx[17] := UDINT_TO_BYTE(SHR(nStartAddr, 16) AND 16#FF);

        // 1.11. Device Code (M=0x90, D=0xA8, ...)
        aTx[18] := TO_BYTE(eDevice);

        // 1.12. Number of Device Points (2 bytes: LSB -> MSB)
        aTx[19] := UINT_TO_BYTE(nPoints AND 16#FF);
        aTx[20] := UINT_TO_BYTE(SHR(nPoints, 8) AND 16#FF);

        bBusy  := TRUE;
        bOwnsSession := TRUE;
        nRxCount := 0;
        nExpectedFrame := 0;
        nState := 10;
    END_IF;
END_IF;


// ================================================================
// MÁY TRẠNG THÁI GIAO TIẾP SOCKET
// ================================================================
CASE nState OF

    10: // PHÁT LỆNH GỬI KHUNG REQUEST
        fbSend(
            sSrvNetId := '',
            hSocket   := stSession.hSocket,
            cbLen     := 21,
            pSrc      := ADR(aTx),
            bExecute  := TRUE,
            tTimeout  := T#3S
        );

        nState := 11;


    11: // CHỜ GỬI XONG
        fbSend(
            sSrvNetId := '',
            hSocket   := stSession.hSocket,
            cbLen     := 21,
            pSrc      := ADR(aTx),
            bExecute  := FALSE,
            tTimeout  := T#3S
        );

        IF NOT fbSend.bBusy THEN
            IF fbSend.bError THEN
                bError   := TRUE;
                nErrorID := fbSend.nErrId;
                stSession.bConnected := FALSE;
                bBusy    := FALSE;
                nState   := 0;
            ELSE
                nState := 20;
            END_IF;
        END_IF;


    20: // PHÁT LỆNH NHẬN RESPONSE
        fbReceive(
            sSrvNetId := '',
            hSocket   := stSession.hSocket,
            cbLen     := SIZEOF(aRx) - nRxCount,
            pDest     := ADR(aRx[nRxCount]),
            bExecute  := TRUE,
            tTimeout  := T#3S
        );

        nState := 21;


    21: // CHỜ PLC-Q TRẢ RESPONSE (Polled receive với timeout 2 giây)
        fbReceive(
            sSrvNetId := '',
            hSocket   := stSession.hSocket,
            cbLen     := SIZEOF(aRx) - nRxCount,
            pDest     := ADR(aRx[nRxCount]),
            bExecute  := FALSE,
            tTimeout  := T#3S
        );

        IF NOT fbReceive.bBusy THEN
            IF fbReceive.bError THEN
                bError   := TRUE;
                nErrorID := fbReceive.nErrId;
                stSession.bConnected := FALSE;
                bBusy    := FALSE;
                nState   := 0;

